      W_g[13,34] := -0.05300187;
      W_g[13,35] := -0.05293896;
      W_g[13,36] := 0.09086524;
      W_g[13,37] := 0.02082952;
      W_g[13,38] := -0.06235110;
      W_g[13,39] := 0.00900952;
      W_g[14,0] := -0.11502921;
      W_g[14,1] := -0.07562436;
      W_g[14,2] := 0.11307055;
      W_g[14,3] := -0.26701322;
      W_g[14,4] := -0.58367014;
      W_g[14,5] := -0.36228108;
      W_g[14,6] := -0.67209059;
      W_g[14,7] := -0.12579566;
      W_g[14,8] := 0.09378675;
      W_g[14,9] := 0.05906596;
      W_g[14,10] := 0.16357109;
      W_g[14,11] := -0.32748589;
      W_g[14,12] := 0.37227204;
      W_g[14,13] := -0.05649122;
      W_g[14,14] := -0.05130398;
      W_g[14,15] := 0.17849237;
      W_g[14,16] := -0.01951551;
      W_g[14,17] := -0.03428079;
      W_g[14,18] := 0.00277206;
      W_g[14,19] := -0.03570505;
      W_g[14,20] := -0.25614583;
      W_g[14,21] := 0.05955129;
      W_g[14,22] := 0.00051241;
      W_g[14,23] := -0.01442853;
      W_g[14,24] := 0.26009023;
      W_g[14,25] := 0.06896590;
      W_g[14,26] := -0.08565364;
      W_g[14,27] := -0.03922650;
      W_g[14,28] := 0.49202508;
      W_g[14,29] := -0.49808294;
      W_g[14,30] := 0.13317353;
      W_g[14,31] := -0.11772110;
      W_g[14,32] := -0.11562508;
      W_g[14,33] := -0.08904682;
      W_g[14,34] := -0.06742100;
      W_g[14,35] := 0.08811268;
      W_g[14,36] := 0.09177279;
      W_g[14,37] := 0.04189566;
      W_g[14,38] := -0.02056031;
      W_g[14,39] := 0.12051180;
      W_g[15,0] := 0.15540718;
      W_g[15,1] := 0.07573265;
      W_g[15,2] := -0.25493059;
      W_g[15,3] := -0.14080612;
      W_g[15,4] := -0.16169477;
      W_g[15,5] := -0.00757927;
      W_g[15,6] := 0.08066899;
      W_g[15,7] := 0.01200249;
      W_g[15,8] := 0.03001926;
      W_g[15,9] := 0.11639266;
      W_g[15,10] := 0.07306892;
      W_g[15,11] := 0.28355977;
      W_g[15,12] := 0.48124212;
      W_g[15,13] := -0.12040935;
      W_g[15,14] := 0.02596140;
      W_g[15,15] := -0.21398795;
      W_g[15,16] := -0.09279459;
      W_g[15,17] := 0.00674920;
      W_g[15,18] := 0.21276073;
      W_g[15,19] := -0.03845788;
      W_g[15,20] := -0.04765760;
      W_g[15,21] := 0.01264688;
      W_g[15,22] := -0.01257103;
      W_g[15,23] := -0.06903563;
      W_g[15,24] := -0.15318221;
      W_g[15,25] := -0.25217903;
      W_g[15,26] := -0.03703345;
      W_g[15,27] := -0.10722972;
      W_g[15,28] := 0.05285160;
      W_g[15,29] := 0.08407086;
      W_g[15,30] := -0.01538745;
      W_g[15,31] := 0.00114667;
      W_g[15,32] := -0.07507251;
      W_g[15,33] := -0.06782222;
      W_g[15,34] := -0.36006817;
      W_g[15,35] := -0.05444269;
      W_g[15,36] := -0.01375175;
      W_g[15,37] := -0.02703385;
      W_g[15,38] := 0.45141658;
      W_g[15,39] := -0.03576548;
      W_g[16,0] := -0.01573141;
      W_g[16,1] := -0.01249725;
      W_g[16,2] := -0.01918053;
      W_g[16,3] := -0.32394302;
      W_g[16,4] := -0.06679904;
      W_g[16,5] := 0.09351813;
      W_g[16,6] := -0.03767738;
      W_g[16,7] := 0.01552502;
      W_g[16,8] := 0.02639228;
      W_g[16,9] := 0.27829525;
      W_g[16,10] := 0.01795475;
      W_g[16,11] := 0.61483020;
      W_g[16,12] := -0.23530579;
      W_g[16,13] := -0.10427370;
      W_g[16,14] := -0.00830992;
      W_g[16,15] := -0.04126130;
      W_g[16,16] := 0.02147032;
      W_g[16,17] := 0.22274575;
      W_g[16,18] := -0.05346655;
      W_g[16,19] := 0.59863454;
      W_g[16,20] := 0.02781765;
      W_g[16,21] := 0.03784034;
      W_g[16,22] := -0.01627534;
      W_g[16,23] := -0.09212849;
      W_g[16,24] := 0.20988049;
      W_g[16,25] := 0.11980043;
      W_g[16,26] := -0.06347527;
      W_g[16,27] := 0.03875433;
      W_g[16,28] := -0.00814277;
      W_g[16,29] := -0.01749807;
      W_g[16,30] := -0.11471809;
      W_g[16,31] := 0.03057062;
      W_g[16,32] := 0.05926932;
      W_g[16,33] := 0.07752163;
      W_g[16,34] := 0.30541685;
      W_g[16,35] := 0.08390119;
      W_g[16,36] := 0.01792176;
      W_g[16,37] := 0.07683819;
      W_g[16,38] := -0.12264256;
      W_g[16,39] := -0.29801413;
      W_g[17,0] := -0.20019235;
      W_g[17,1] := 0.08634444;
      W_g[17,2] := 0.35990810;
      W_g[17,3] := -0.54319084;
      W_g[17,4] := 0.10491174;
      W_g[17,5] := -0.24461722;
      W_g[17,6] := 0.00542844;
      W_g[17,7] := -0.00443292;
      W_g[17,8] := -0.13760753;
      W_g[17,9] := 0.17179628;
      W_g[17,10] := 0.57468456;
      W_g[17,11] := 0.84765750;
      W_g[17,12] := -0.84660238;
      W_g[17,13] := -0.02827467;
      W_g[17,14] := 0.09285270;
      W_g[17,15] := 0.00605520;
      W_g[17,16] := -0.23755617;
      W_g[17,17] := 0.01386433;
      W_g[17,18] := 0.00373611;
      W_g[17,19] := 0.64604604;
      W_g[17,20] := -0.30180034;
      W_g[17,21] := -0.71723890;
      W_g[17,22] := -0.23780504;
      W_g[17,23] := 0.04141965;
      W_g[17,24] := -0.74509096;
      W_g[17,25] := -0.75259161;
      W_g[17,26] := 0.24358149;
      W_g[17,27] := 0.62698990;
      W_g[17,28] := -0.24088508;
      W_g[17,29] := 0.06953070;
      W_g[17,30] := -0.33534220;
      W_g[17,31] := -0.02631341;
      W_g[17,32] := -0.30826521;
      W_g[17,33] := -0.45180380;
      W_g[17,34] := -0.90610892;
      W_g[17,35] := -0.06815604;
      W_g[17,36] := -0.14631121;
      W_g[17,37] := 0.17388295;
      W_g[17,38] := 0.13864316;
      W_g[17,39] := 0.17807765;
      W_g[18,0] := -0.46607670;
      W_g[18,1] := 0.10845635;
      W_g[18,2] := 0.22516194;
      W_g[18,3] := 0.30607522;
      W_g[18,4] := -0.15093884;
      W_g[18,5] := 0.01696070;
      W_g[18,6] := 0.16042185;
      W_g[18,7] := -0.10679442;
      W_g[18,8] := 0.20514138;
      W_g[18,9] := -0.13397862;
      W_g[18,10] := 0.02242056;
      W_g[18,11] := -0.19990624;
      W_g[18,12] := 0.38241696;
      W_g[18,13] := -0.01298471;
      W_g[18,14] := -0.00218331;
      W_g[18,15] := -0.04433896;
      W_g[18,16] := -0.26164895;
      W_g[18,17] := 0.05559360;
      W_g[18,18] := -0.06075819;
      W_g[18,19] := -0.05308994;
      W_g[18,20] := -0.13432083;
      W_g[18,21] := -0.33185339;
      W_g[18,22] := -0.08431048;
      W_g[18,23] := -0.16004905;
      W_g[18,24] := -0.36850065;
      W_g[18,25] := -0.04567018;
      W_g[18,26] := -0.34792730;
      W_g[18,27] := -0.06563149;
      W_g[18,28] := 0.04670760;
      W_g[18,29] := 0.06350503;
      W_g[18,30] := -0.07850740;
      W_g[18,31] := 0.16866533;
      W_g[18,32] := 0.02046569;
      W_g[18,33] := 0.05549860;
      W_g[18,34] := 0.01890240;
      W_g[18,35] := -0.02811935;
      W_g[18,36] := 0.03381456;
      W_g[18,37] := 0.11580943;
      W_g[18,38] := -0.11624962;
      W_g[18,39] := -0.03905239;
      W_g[19,0] := 0.01773376;
      W_g[19,1] := -0.05072702;
      W_g[19,2] := -0.00225121;
      W_g[19,3] := -0.01785041;
      W_g[19,4] := 0.04858205;
      W_g[19,5] := -0.01839915;
      W_g[19,6] := -0.04408873;
      W_g[19,7] := -0.01353623;
      W_g[19,8] := -0.00090088;
      W_g[19,9] := -0.00116132;
      W_g[19,10] := 0.00882178;
      W_g[19,11] := -0.03854829;
      W_g[19,12] := 0.03738030;
      W_g[19,13] := -0.01948604;
      W_g[19,14] := -0.45808697;
      W_g[19,15] := -0.26110804;
      W_g[19,16] := 0.00333187;
      W_g[19,17] := -0.25176817;
      W_g[19,18] := 0.08445162;
      W_g[19,19] := 0.26523203;
      W_g[19,20] := -0.05709776;
      W_g[19,21] := -0.05241840;
      W_g[19,22] := 0.01751016;
      W_g[19,23] := -0.00974986;
      W_g[19,24] := 0.27344036;
      W_g[19,25] := 0.32422283;
      W_g[19,26] := -0.04881701;
      W_g[19,27] := -0.02297378;
      W_g[19,28] := -0.06826914;
      W_g[19,29] := -0.11992263;
      W_g[19,30] := 0.01903425;
      W_g[19,31] := 0.02200578;
      W_g[19,32] := -0.04815840;
      W_g[19,33] := -0.11233919;
      W_g[19,34] := -0.23930897;
      W_g[19,35] := 0.02726550;
      W_g[19,36] := -0.00201288;
      W_g[19,37] := 0.05262006;
      W_g[19,38] := -0.04631574;
      W_g[19,39] := -0.25027138;
      W_g[20,0] := -0.17776611;
      W_g[20,1] := -0.49992636;
      W_g[20,2] := 0.03143674;
      W_g[20,3] := 0.15612000;
      W_g[20,4] := -0.50436848;
      W_g[20,5] := 0.02739897;
      W_g[20,6] := -0.10362915;
      W_g[20,7] := 0.35108495;
      W_g[20,8] := 0.19622006;
      W_g[20,9] := 0.38027030;
      W_g[20,10] := -0.53794569;
      W_g[20,11] := 0.05582263;
      W_g[20,12] := -0.17187732;
      W_g[20,13] := -0.14350507;
      W_g[20,14] := 0.04435784;
      W_g[20,15] := -0.00301744;
      W_g[20,16] := 0.05593058;
      W_g[20,17] := 0.00574902;
      W_g[20,18] := 0.02816820;
      W_g[20,19] := -0.00896498;
      W_g[20,20] := -0.27302650;
      W_g[20,21] := -0.10916554;
      W_g[20,22] := 0.07598325;
      W_g[20,23] := 0.07597133;
      W_g[20,24] := -0.20816125;
      W_g[20,25] := -0.00556583;
      W_g[20,26] := 0.15926160;
      W_g[20,27] := 0.04909170;
      W_g[20,28] := -0.30622017;
      W_g[20,29] := 0.16263185;
      W_g[20,30] := 0.06980544;
      W_g[20,31] := 0.18102454;
      W_g[20,32] := 0.01593671;
      W_g[20,33] := -0.04853294;
      W_g[20,34] := -0.09243315;
      W_g[20,35] := 0.03795157;
      W_g[20,36] := -0.01642190;
      W_g[20,37] := 0.06450415;
      W_g[20,38] := -0.01715147;
      W_g[20,39] := -0.05797761;
      W_g[21,0] := 0.04719520;
      W_g[21,1] := 0.01569074;
      W_g[21,2] := -0.00857600;
      W_g[21,3] := 0.36854166;
      W_g[21,4] := -0.29962948;
      W_g[21,5] := 0.11101421;
      W_g[21,6] := -0.14704654;
      W_g[21,7] := -0.25060529;
      W_g[21,8] := 0.03979661;
      W_g[21,9] := -0.37424278;
      W_g[21,10] := 0.33715650;
      W_g[21,11] := 0.20566781;
      W_g[21,12] := -0.55089366;
      W_g[21,13] := -0.34874550;
      W_g[21,14] := -0.00000745;
      W_g[21,15] := 0.11779826;
      W_g[21,16] := -0.01198818;
      W_g[21,17] := -0.09557019;
      W_g[21,18] := -0.38575107;
      W_g[21,19] := 0.10345905;
      W_g[21,20] := 0.17967871;
      W_g[21,21] := -0.02546586;
      W_g[21,22] := 0.02202458;
      W_g[21,23] := -0.47533408;
      W_g[21,24] := -0.07804859;
      W_g[21,25] := -0.20474817;
      W_g[21,26] := 0.09593988;
      W_g[21,27] := -0.20002005;
      W_g[21,28] := 0.14636038;
      W_g[21,29] := 0.27730727;
      W_g[21,30] := 0.03117772;
      W_g[21,31] := 0.06990665;
      W_g[21,32] := 0.05139569;
      W_g[21,33] := 0.08534111;
      W_g[21,34] := 0.34672982;
      W_g[21,35] := 0.01232039;
      W_g[21,36] := -0.05206082;
      W_g[21,37] := -0.01625307;
      W_g[21,38] := 0.20143867;
      W_g[21,39] := -0.10067950;
      W_g[22,0] := 0.11665134;
      W_g[22,1] := 0.10529415;
      W_g[22,2] := 0.22086281;
      W_g[22,3] := -0.12558044;
      W_g[22,4] := -0.00237558;
      W_g[22,5] := 0.19240804;
      W_g[22,6] := -0.24772990;
      W_g[22,7] := 0.08354132;
      W_g[22,8] := -0.20447712;
      W_g[22,9] := 0.03358927;
      W_g[22,10] := -0.15093991;
      W_g[22,11] := -0.03152904;
      W_g[22,12] := 0.23958053;
      W_g[22,13] := -0.10689051;
      W_g[22,14] := 0.14513183;
      W_g[22,15] := 0.20699252;
      W_g[22,16] := -0.00007249;
      W_g[22,17] := 0.01122855;
      W_g[22,18] := -0.00866538;
      W_g[22,19] := 0.10550721;
      W_g[22,20] := -0.14577182;
      W_g[22,21] := 0.25070757;
      W_g[22,22] := 0.07765597;
      W_g[22,23] := 0.12089684;
      W_g[22,24] := 0.42342681;
      W_g[22,25] := 0.12979737;
      W_g[22,26] := 0.16623591;
      W_g[22,27] := -0.09820254;
      W_g[22,28] := 0.03250218;
      W_g[22,29] := 0.11340379;
      W_g[22,30] := 0.08371338;
      W_g[22,31] := 0.10858538;
      W_g[22,32] := -0.09717516;
      W_g[22,33] := -0.05043048;
      W_g[22,34] := -0.12874730;
      W_g[22,35] := -0.16679265;
      W_g[22,36] := 0.06777173;
      W_g[22,37] := -0.19872338;
      W_g[22,38] := -0.09894791;
      W_g[22,39] := -0.29871914;
      W_g[23,0] := -0.07641292;
      W_g[23,1] := -0.00534786;
      W_g[23,2] := 0.20778368;
      W_g[23,3] := 0.22361241;
      W_g[23,4] := 0.03807362;
      W_g[23,5] := -0.02697703;
      W_g[23,6] := -0.13366827;
      W_g[23,7] := -0.03372496;
      W_g[23,8] := -0.11303925;
      W_g[23,9] := -0.14616819;
      W_g[23,10] := 0.00094925;
      W_g[23,11] := 0.17858963;
      W_g[23,12] := -0.02489791;
      W_g[23,13] := -0.03910236;
      W_g[23,14] := -0.02416698;
      W_g[23,15] := -0.25673768;
      W_g[23,16] := 0.30395365;
      W_g[23,17] := -0.01390388;
      W_g[23,18] := 0.00377696;
      W_g[23,19] := 0.08999401;
      W_g[23,20] := -0.40618902;
      W_g[23,21] := -0.18011197;
      W_g[23,22] := -0.10348500;
      W_g[23,23] := 0.01184078;
      W_g[23,24] := -0.60941619;
      W_g[23,25] := -0.17570031;
      W_g[23,26] := 0.09114521;
      W_g[23,27] := 0.07809471;
      W_g[23,28] := -0.03781823;
      W_g[23,29] := -0.02985572;
      W_g[23,30] := -0.10175200;
      W_g[23,31] := 0.07091261;
      W_g[23,32] := 0.00975894;
      W_g[23,33] := 0.07413130;
      W_g[23,34] := 0.04860087;
      W_g[23,35] := -0.06112134;
      W_g[23,36] := -0.01834961;
      W_g[23,37] := -0.06767160;
      W_g[23,38] := 0.04615815;
      W_g[23,39] := 0.03219241;
      W_g[24,0] := 0.14109130;
      W_g[24,1] := 0.23656085;
      W_g[24,2] := -0.05220996;
      W_g[24,3] := -0.08191337;
      W_g[24,4] := -0.59643692;
      W_g[24,5] := -0.08740985;
      W_g[24,6] := 0.51112539;
      W_g[24,7] := -0.08679886;
      W_g[24,8] := -0.03170026;
      W_g[24,9] := -0.04040290;
      W_g[24,10] := 0.42674446;
      W_g[24,11] := 0.22892350;
      W_g[24,12] := 0.06517982;
      W_g[24,13] := -0.07052775;
      W_g[24,14] := 0.00610844;
      W_g[24,15] := -0.14473575;
      W_g[24,16] := 0.11628936;
      W_g[24,17] := 0.00950560;
      W_g[24,18] := -0.05220868;
      W_g[24,19] := -0.21057445;
      W_g[24,20] := 0.15953180;
      W_g[24,21] := 0.03443460;
      W_g[24,22] := 0.02498991;
      W_g[24,23] := 0.15479933;
      W_g[24,24] := 0.31532544;
      W_g[24,25] := -0.07248386;
      W_g[24,26] := 0.22804081;
      W_g[24,27] := -0.23870072;
      W_g[24,28] := 0.07509667;
      W_g[24,29] := -0.04223498;
      W_g[24,30] := 0.02754644;
      W_g[24,31] := 0.04945280;
      W_g[24,32] := -0.12835518;
      W_g[24,33] := -0.16013861;
      W_g[24,34] := -0.20117347;
      W_g[24,35] := -0.09332737;
      W_g[24,36] := -0.27658218;
      W_g[24,37] := -0.14927265;
      W_g[24,38] := -0.28982732;
      W_g[24,39] := 0.01216547;
      W_g[25,0] := 0.00249727;
      W_g[25,1] := 0.02321395;
      W_g[25,2] := 0.03579676;
      W_g[25,3] := -0.32325658;
      W_g[25,4] := 0.07457885;
      W_g[25,5] := 0.01599968;
      W_g[25,6] := -0.19957243;
      W_g[25,7] := 0.12909044;
      W_g[25,8] := 0.00623424;
      W_g[25,9] := 0.26816839;
      W_g[25,10] := -0.23799382;
      W_g[25,11] := -0.18556090;
      W_g[25,12] := -0.03897551;
      W_g[25,13] := -0.07030228;
      W_g[25,14] := -0.06287792;
      W_g[25,15] := 0.17744720;
      W_g[25,16] := -0.03842967;
      W_g[25,17] := -0.06559484;
      W_g[25,18] := 0.02993315;
      W_g[25,19] := 0.08945196;
      W_g[25,20] := -0.00580116;
      W_g[25,21] := -0.02753790;
      W_g[25,22] := -0.02607165;
      W_g[25,23] := -0.00466925;
      W_g[25,24] := -0.84821171;
      W_g[25,25] := 0.23694646;
      W_g[25,26] := -0.14543480;
      W_g[25,27] := -0.15780894;
      W_g[25,28] := -0.27692312;
      W_g[25,29] := -0.04585484;
      W_g[25,30] := -0.03756009;
      W_g[25,31] := -0.08991528;
      W_g[25,32] := 0.00971850;
      W_g[25,33] := 0.08656777;
      W_g[25,34] := 0.12360313;
      W_g[25,35] := -0.08704287;
      W_g[25,36] := -0.50061452;
      W_g[25,37] := 0.06715164;
      W_g[25,38] := 0.03072628;
      W_g[25,39] := -0.05923472;
      W_g[26,0] := 0.19895676;
      W_g[26,1] := 0.01795273;
      W_g[26,2] := -0.08949947;
      W_g[26,3] := -0.06816271;
      W_g[26,4] := -0.12828159;
      W_g[26,5] := 0.00080027;
      W_g[26,6] := 0.16275345;
      W_g[26,7] := 0.14247812;
      W_g[26,8] := -0.05336298;
      W_g[26,9] := 0.16001105;
      W_g[26,10] := -0.00170321;
      W_g[26,11] := -0.10854331;
      W_g[26,12] := 0.11391646;
      W_g[26,13] := 0.31833315;
      W_g[26,14] := -0.00052231;
      W_g[26,15] := 0.04305906;
      W_g[26,16] := -0.00767927;
      W_g[26,17] := -0.03174791;
      W_g[26,18] := -1.20069015;
      W_g[26,19] := 0.08255526;
      W_g[26,20] := -0.47470504;
      W_g[26,21] := 0.21856050;
      W_g[26,22] := 0.04315476;
      W_g[26,23] := 0.15731587;
      W_g[26,24] := -0.16662689;
      W_g[26,25] := -0.36638814;
      W_g[26,26] := -0.28305781;
      W_g[26,27] := -0.09379881;
      W_g[26,28] := -0.24579851;
      W_g[26,29] := 0.01016386;
      W_g[26,30] := 0.01751088;
      W_g[26,31] := 0.15965039;
      W_g[26,32] := 0.00510592;
      W_g[26,33] := 0.09451680;
      W_g[26,34] := 0.02374958;
      W_g[26,35] := -0.10228859;
      W_g[26,36] := 0.04589900;
      W_g[26,37] := -0.01942009;
      W_g[26,38] := 0.15447062;
      W_g[26,39] := -0.00123656;
      W_g[27,0] := -0.14282966;
      W_g[27,1] := 0.03789151;
      W_g[27,2] := 0.02735430;
      W_g[27,3] := -0.02859589;
      W_g[27,4] := 0.11969381;
      W_g[27,5] := -0.08108735;
      W_g[27,6] := -0.48059788;
      W_g[27,7] := 0.11670560;
      W_g[27,8] := 0.02436283;
      W_g[27,9] := 0.15240525;
      W_g[27,10] := 0.60784400;
      W_g[27,11] := 0.16673699;
      W_g[27,12] := -0.11131126;
      W_g[27,13] := 0.39158168;
      W_g[27,14] := -0.01387984;
      W_g[27,15] := 0.03263223;
      W_g[27,16] := 0.07995110;
      W_g[27,17] := -0.01656702;
      W_g[27,18] := 0.16666247;
      W_g[27,19] := -0.07363571;
      W_g[27,20] := -0.26380217;
      W_g[27,21] := 0.36762938;
      W_g[27,22] := 0.10293096;
      W_g[27,23] := -0.21954748;
      W_g[27,24] := -0.19905801;
      W_g[27,25] := 0.00590560;
      W_g[27,26] := -0.07474038;
      W_g[27,27] := -0.00682373;
      W_g[27,28] := 0.00600550;
      W_g[27,29] := 0.52201474;
      W_g[27,30] := 0.10763236;
      W_g[27,31] := 0.20513408;
      W_g[27,32] := 0.08530629;
      W_g[27,33] := 0.18354966;
      W_g[27,34] := 0.20833531;
      W_g[27,35] := -0.02688346;
      W_g[27,36] := -0.05211073;
      W_g[27,37] := -0.10546255;
      W_g[27,38] := -0.16810939;
      W_g[27,39] := 0.04055268;
      W_g[28,0] := -0.12039233;
      W_g[28,1] := 0.03123983;
      W_g[28,2] := -0.28947538;
      W_g[28,3] := -0.24017365;
      W_g[28,4] := 0.29521075;
      W_g[28,5] := 0.08690419;
      W_g[28,6] := 0.01901748;
      W_g[28,7] := -0.23417597;
      W_g[28,8] := 0.43286511;
      W_g[28,9] := 0.02607675;
      W_g[28,10] := 0.19849846;
      W_g[28,11] := -0.06265938;
      W_g[28,12] := 0.09416307;
      W_g[28,13] := -0.05105516;
      W_g[28,14] := -0.01597860;
      W_g[28,15] := 0.14792809;
      W_g[28,16] := 0.14414477;
      W_g[28,17] := -0.02288275;
      W_g[28,18] := -0.03377746;
      W_g[28,19] := -0.15792006;
      W_g[28,20] := -0.21533181;
      W_g[28,21] := 0.08094171;
      W_g[28,22] := 0.00793070;
      W_g[28,23] := 0.03326877;
      W_g[28,24] := 0.04408788;
      W_g[28,25] := -0.11347675;
      W_g[28,26] := 0.14422546;
      W_g[28,27] := 0.19584695;
      W_g[28,28] := -0.13756958;
      W_g[28,29] := -0.12223729;
      W_g[28,30] := 0.02110463;
      W_g[28,31] := 0.03519979;
      W_g[28,32] := -0.05562153;
      W_g[28,33] := -0.06591920;
      W_g[28,34] := 0.04866378;
      W_g[28,35] := -0.09032071;
      W_g[28,36] := 0.03939996;
      W_g[28,37] := -0.08595932;
      W_g[28,38] := 0.01556356;
      W_g[28,39] := -0.17334549;
      W_g[29,0] := -0.01603005;
      W_g[29,1] := 0.00894765;
      W_g[29,2] := 0.04728428;
      W_g[29,3] := 0.13398947;
      W_g[29,4] := -0.08206625;
      W_g[29,5] := 0.43515241;
      W_g[29,6] := -0.08524376;
      W_g[29,7] := 0.12636763;
      W_g[29,8] := -0.07064829;
      W_g[29,9] := 0.02922662;
      W_g[29,10] := 0.16617142;
      W_g[29,11] := -0.03181689;
      W_g[29,12] := -0.18755385;
      W_g[29,13] := 0.04736114;
      W_g[29,14] := 0.00172536;
      W_g[29,15] := 0.02388163;
      W_g[29,16] := -0.00605842;
      W_g[29,17] := -0.00226685;
      W_g[29,18] := 0.18417786;
      W_g[29,19] := 0.02931385;
      W_g[29,20] := -0.10084365;
      W_g[29,21] := -0.03299641;
      W_g[29,22] := -0.00275616;
      W_g[29,23] := 0.02141913;
      W_g[29,24] := 0.00477037;
      W_g[29,25] := 0.05081034;
      W_g[29,26] := -0.19006838;
      W_g[29,27] := -0.14232871;
      W_g[29,28] := 0.06605857;
      W_g[29,29] := -0.26251897;
      W_g[29,30] := -0.00548652;
      W_g[29,31] := 0.03245487;
      W_g[29,32] := -0.05614575;
      W_g[29,33] := -0.08672421;
      W_g[29,34] := -0.19275941;
      W_g[29,35] := -0.02231585;
      W_g[29,36] := 0.00673404;
      W_g[29,37] := -0.02077745;
      W_g[29,38] := 0.02013531;
      W_g[29,39] := 0.21206558;
      W_g[30,0] := 0.06752372;
      W_g[30,1] := 0.04914160;
      W_g[30,2] := 0.03581399;
      W_g[30,3] := 0.55463815;
      W_g[30,4] := 0.19955039;
      W_g[30,5] := -0.29638356;
      W_g[30,6] := 0.61677969;
      W_g[30,7] := -0.08204620;
      W_g[30,8] := -0.02945163;
      W_g[30,9] := -0.33782583;
      W_g[30,10] := 0.03250416;
      W_g[30,11] := 0.32107306;
      W_g[30,12] := 0.06659118;
      W_g[30,13] := 0.29332143;
      W_g[30,14] := -0.02582538;
      W_g[30,15] := 0.62199312;
      W_g[30,16] := 0.28212488;
      W_g[30,17] := -0.23582231;
      W_g[30,18] := 0.33779177;
      W_g[30,19] := 0.50508004;
      W_g[30,20] := -0.04146927;
      W_g[30,21] := 0.00146027;
      W_g[30,22] := 0.10298456;
      W_g[30,23] := -0.13510256;
      W_g[30,24] := 0.08098176;
      W_g[30,25] := -0.07603540;
      W_g[30,26] := 0.11315724;
      W_g[30,27] := 0.12087354;
      W_g[30,28] := -0.23194072;
      W_g[30,29] := 0.06172852;
      W_g[30,30] := 0.06911052;
      W_g[30,31] := 0.33844078;
      W_g[30,32] := 0.07554214;
      W_g[30,33] := 0.01718852;
      W_g[30,34] := -0.07873586;
      W_g[30,35] := -0.07006503;
      W_g[30,36] := 0.00541107;
      W_g[30,37] := -0.08336300;
      W_g[30,38] := 0.02301235;
      W_g[30,39] := 0.23563193;
      W_g[31,0] := 0.18860947;
      W_g[31,1] := -0.02123935;
      W_g[31,2] := -0.26690537;
      W_g[31,3] := 0.12378932;
      W_g[31,4] := 0.09037927;
      W_g[31,5] := -0.03088225;
      W_g[31,6] := -0.17878367;
      W_g[31,7] := 0.02112429;
      W_g[31,8] := 0.03763676;
      W_g[31,9] := -0.02504454;
      W_g[31,10] := -0.01659736;
      W_g[31,11] := 0.16001292;
      W_g[31,12] := -0.06862063;
      W_g[31,13] := -0.08124028;
      W_g[31,14] := -0.00468529;
      W_g[31,15] := -0.14859970;
      W_g[31,16] := -0.30615747;
      W_g[31,17] := -0.02353984;
      W_g[31,18] := 0.01195374;
      W_g[31,19] := 0.04420421;
      W_g[31,20] := -0.08521901;
      W_g[31,21] := 0.06032958;
      W_g[31,22] := 0.01825500;
      W_g[31,23] := 0.05283485;
      W_g[31,24] := -0.25803921;
      W_g[31,25] := 0.03302622;
      W_g[31,26] := 0.16146830;
      W_g[31,27] := 0.17279540;
      W_g[31,28] := 0.01809685;
      W_g[31,29] := 0.02630481;
      W_g[31,30] := 0.03338469;
      W_g[31,31] := 0.45954949;
      W_g[31,32] := -0.04697010;
      W_g[31,33] := 0.03801997;
      W_g[31,34] := 0.22326140;
      W_g[31,35] := -0.18952455;
      W_g[31,36] := 0.00136513;
      W_g[31,37] := -0.27123162;
      W_g[31,38] := -0.07247190;
      W_g[31,39] := 0.23167513;
      W_o[0,0] := 0.42249125;
      W_o[0,1] := -0.64850706;
      W_o[0,2] := -0.08193821;
      W_o[0,3] := -0.33892727;
      W_o[0,4] := 0.05321682;
      W_o[0,5] := 0.11530717;
      W_o[0,6] := 0.32608813;
      W_o[0,7] := -0.13539509;
      W_o[0,8] := 0.20117587;
      W_o[0,9] := -0.31878343;
      W_o[0,10] := -0.17219098;
      W_o[0,11] := 0.14882079;
      W_o[0,12] := 0.11313346;
      W_o[0,13] := -0.10760950;
      W_o[0,14] := 0.01743469;
      W_o[0,15] := 0.01349122;
      W_o[0,16] := -0.01363511;
      W_o[0,17] := -0.00418937;
      W_o[0,18] := -0.08654208;
      W_o[0,19] := 0.01018774;
      W_o[0,20] := 0.37044030;
      W_o[0,21] := 0.87406963;
      W_o[0,22] := 0.05330493;
      W_o[0,23] := -0.60551524;
      W_o[0,24] := 0.00528000;
      W_o[0,25] := 0.00492091;
      W_o[0,26] := -0.73618817;
      W_o[0,27] := 0.86269325;
      W_o[0,28] := 0.67136478;
      W_o[0,29] := -0.14723247;
      W_o[0,30] := -0.17640491;
      W_o[0,31] := 0.00200789;
      W_o[0,32] := -0.11784527;
      W_o[0,33] := 0.32575944;
      W_o[0,34] := 0.11160263;
      W_o[0,35] := -0.05652209;
      W_o[0,36] := 0.04402122;
      W_o[0,37] := 0.08225929;
      W_o[0,38] := 0.20138605;
      W_o[0,39] := -0.07881875;
      W_o[1,0] := -1.27534890;
      W_o[1,1] := -0.27924889;
      W_o[1,2] := -0.75771481;
      W_o[1,3] := -0.18380418;
      W_o[1,4] := -0.39482769;
      W_o[1,5] := 0.10104305;
      W_o[1,6] := -0.34825188;
      W_o[1,7] := -0.63163066;
      W_o[1,8] := -1.08178067;
      W_o[1,9] := -0.97093791;
      W_o[1,10] := -0.20904520;
      W_o[1,11] := -0.29529026;
      W_o[1,12] := -0.14393961;
      W_o[1,13] := -0.01520389;
      W_o[1,14] := 0.00541295;
      W_o[1,15] := -0.02735653;
      W_o[1,16] := -0.07699423;
      W_o[1,17] := 0.08873669;
      W_o[1,18] := 0.18124166;
      W_o[1,19] := -0.01098941;
      W_o[1,20] := 0.13787243;
      W_o[1,21] := 0.26410136;
      W_o[1,22] := 0.06537609;
      W_o[1,23] := -0.15175536;
      W_o[1,24] := -0.11301857;
      W_o[1,25] := -0.10047740;
      W_o[1,26] := 0.11024941;
      W_o[1,27] := 0.24368817;
      W_o[1,28] := 0.59257942;
      W_o[1,29] := 0.02251752;
      W_o[1,30] := 0.20542605;
      W_o[1,31] := 0.05349508;
      W_o[1,32] := 0.07199062;
      W_o[1,33] := 0.06075877;
      W_o[1,34] := 0.17365526;
      W_o[1,35] := -0.04894430;
      W_o[1,36] := -0.02975028;
      W_o[1,37] := -0.12903002;
      W_o[1,38] := 0.08992038;
      W_o[1,39] := 0.10337646;
      W_o[2,0] := 0.30405313;
      W_o[2,1] := 0.00766394;
      W_o[2,2] := -0.18612629;
      W_o[2,3] := 0.15926282;
      W_o[2,4] := 0.50370109;
      W_o[2,5] := 0.69898289;
      W_o[2,6] := 1.03120697;
      W_o[2,7] := 0.06395171;
      W_o[2,8] := 0.13832410;
      W_o[2,9] := 0.10960636;
      W_o[2,10] := -0.42085138;
      W_o[2,11] := 0.39040789;
      W_o[2,12] := 0.06325981;
      W_o[2,13] := 0.40687191;
      W_o[2,14] := 0.04082680;
      W_o[2,15] := -0.00324509;
      W_o[2,16] := 0.01833900;
      W_o[2,17] := 0.11513314;
      W_o[2,18] := 0.12066066;
      W_o[2,19] := 0.01082493;
      W_o[2,20] := -0.16976321;
      W_o[2,21] := 0.53049803;
      W_o[2,22] := 0.15725319;
      W_o[2,23] := -0.34637845;
      W_o[2,24] := 1.58245826;
      W_o[2,25] := 1.47554839;
      W_o[2,26] := -0.00448998;
      W_o[2,27] := 0.14077175;
      W_o[2,28] := -0.37107602;
      W_o[2,29] := 0.02695022;
      W_o[2,30] := 0.19601339;
      W_o[2,31] := 0.17389217;
      W_o[2,32] := 0.14344938;
      W_o[2,33] := 0.81406116;
      W_o[2,34] := 1.72799015;
      W_o[2,35] := -0.12091801;
      W_o[2,36] := 0.16224357;
      W_o[2,37] := -0.33939198;
      W_o[2,38] := 0.05670876;
      W_o[2,39] := 0.09963638;
      W_o[3,0] := -0.26549935;
      W_o[3,1] := -0.11039463;
      W_o[3,2] := -0.37164780;
      W_o[3,3] := 0.15892562;
      W_o[3,4] := -0.06230325;
      W_o[3,5] := -0.37457275;
      W_o[3,6] := 0.24259707;
      W_o[3,7] := 0.37691608;
      W_o[3,8] := -0.42493910;
      W_o[3,9] := 0.27702668;
      W_o[3,10] := 0.36755127;
      W_o[3,11] := -0.49238053;
      W_o[3,12] := -0.28828865;
      W_o[3,13] := -0.19150881;
      W_o[3,14] := -0.67414224;
      W_o[3,15] := -0.02529657;
      W_o[3,16] := 0.29622570;
      W_o[3,17] := 0.45850250;
      W_o[3,18] := 0.04778790;
      W_o[3,19] := 0.51993376;
      W_o[3,20] := -0.20207447;
      W_o[3,21] := 0.18979242;
      W_o[3,22] := -0.07848933;
      W_o[3,23] := -0.01705214;
      W_o[3,24] := 0.01806957;
      W_o[3,25] := 0.02297689;
      W_o[3,26] := -0.01870384;
      W_o[3,27] := -0.17662346;
      W_o[3,28] := -0.04692467;
      W_o[3,29] := -0.17209335;
      W_o[3,30] := -0.24459122;
      W_o[3,31] := 0.07113735;
      W_o[3,32] := 0.00606646;
      W_o[3,33] := -0.05090882;
      W_o[3,34] := 0.08984744;
      W_o[3,35] := -0.16125588;
      W_o[3,36] := -0.00926951;
      W_o[3,37] := -0.15794532;
      W_o[3,38] := 0.07680272;
      W_o[3,39] := 1.02147377;
      W_o[4,0] := 0.17977053;
      W_o[4,1] := 0.03995879;
      W_o[4,2] := -0.05187562;
      W_o[4,3] := -0.00068046;
      W_o[4,4] := 0.00082433;
      W_o[4,5] := -0.17477073;
      W_o[4,6] := 0.18298250;
      W_o[4,7] := 0.01242155;
      W_o[4,8] := -0.10564039;
      W_o[4,9] := 0.28895974;
      W_o[4,10] := -0.16322204;
      W_o[4,11] := 0.10945952;
      W_o[4,12] := -0.03262473;
      W_o[4,13] := -0.11646359;
      W_o[4,14] := 0.00214941;
      W_o[4,15] := -0.01470709;
      W_o[4,16] := 0.07081575;
      W_o[4,17] := -0.00195280;
      W_o[4,18] := 0.90504497;
      W_o[4,19] := 0.06995305;
      W_o[4,20] := 0.12764473;
      W_o[4,21] := -0.13823217;
      W_o[4,22] := -0.10447618;
      W_o[4,23] := -0.07500455;
      W_o[4,24] := -0.22946472;
      W_o[4,25] := 0.20651680;
      W_o[4,26] := 0.08378618;
      W_o[4,27] := 0.07185337;
      W_o[4,28] := 0.15295289;
      W_o[4,29] := 0.80911016;
      W_o[4,30] := -0.12649418;
      W_o[4,31] := 0.29769754;
      W_o[4,32] := -0.10073072;
      W_o[4,33] := -0.19524801;
      W_o[4,34] := -0.00692285;
      W_o[4,35] := 0.15373145;
      W_o[4,36] := 0.01237739;
      W_o[4,37] := 0.13210568;
      W_o[4,38] := 0.15424773;
      W_o[4,39] := -0.01015362;
      W_o[5,0] := 0.28912961;
      W_o[5,1] := 2.07105112;
      W_o[5,2] := 0.01252856;
      W_o[5,3] := 0.34673738;
      W_o[5,4] := 0.21192910;
      W_o[5,5] := 0.23409151;
      W_o[5,6] := -0.12695056;
      W_o[5,7] := 0.23784913;
      W_o[5,8] := -0.03728350;
      W_o[5,9] := 0.21514873;
      W_o[5,10] := 0.26284939;
      W_o[5,11] := -0.21792066;
      W_o[5,12] := -0.39795417;
      W_o[5,13] := -0.69216830;
      W_o[5,14] := -0.18849657;
      W_o[5,15] := -0.13393024;
      W_o[5,16] := -0.25170875;
      W_o[5,17] := -0.24293463;
      W_o[5,18] := 0.27309209;
      W_o[5,19] := -0.14950365;
      W_o[5,20] := -0.03219712;
      W_o[5,21] := 0.35288468;
      W_o[5,22] := 0.23942992;
      W_o[5,23] := -0.16948508;
      W_o[5,24] := 1.87266624;
      W_o[5,25] := 1.58824658;
      W_o[5,26] := -0.05295049;
      W_o[5,27] := 0.20530860;
      W_o[5,28] := -0.00417454;
      W_o[5,29] := -0.04709773;
      W_o[5,30] := 0.14920191;
      W_o[5,31] := -0.05560581;
      W_o[5,32] := 0.04669352;
      W_o[5,33] := 0.14553502;
      W_o[5,34] := 0.53250414;
      W_o[5,35] := 0.10384236;
      W_o[5,36] := 0.39177659;
      W_o[5,37] := -0.00503783;
      W_o[5,38] := -0.05498653;
      W_o[5,39] := 0.39836636;
      W_o[6,0] := -0.09602387;
      W_o[6,1] := 0.01318664;
      W_o[6,2] := 0.02895827;
      W_o[6,3] := -0.13262498;
      W_o[6,4] := -0.12622669;
      W_o[6,5] := 0.03745453;
      W_o[6,6] := 0.55729073;
      W_o[6,7] := 0.14179020;
      W_o[6,8] := 0.08813037;
      W_o[6,9] := 0.02709752;
      W_o[6,10] := -0.03546845;
      W_o[6,11] := 0.07040328;
      W_o[6,12] := -0.03574698;
      W_o[6,13] := 0.01986431;
      W_o[6,14] := 0.01404128;
      W_o[6,15] := 0.02171072;
      W_o[6,16] := 0.09358315;
      W_o[6,17] := 0.05428468;
      W_o[6,18] := -0.02667183;
      W_o[6,19] := -0.00128908;
      W_o[6,20] := -1.56595874;
      W_o[6,21] := 0.00646133;
      W_o[6,22] := -0.24436766;
      W_o[6,23] := -0.13901594;
      W_o[6,24] := 0.99376416;
      W_o[6,25] := 0.85211402;
      W_o[6,26] := -0.23664802;
      W_o[6,27] := -0.08933339;
      W_o[6,28] := 0.15226653;
      W_o[6,29] := -0.30946207;
      W_o[6,30] := -0.20975208;
      W_o[6,31] := 0.62505847;
      W_o[6,32] := -0.04092027;
      W_o[6,33] := 0.09183368;
      W_o[6,34] := 0.63159341;
      W_o[6,35] := 0.13661051;
      W_o[6,36] := -0.00265529;
      W_o[6,37] := 0.16893734;
      W_o[6,38] := 0.18080245;
      W_o[6,39] := 0.49472585;
      W_o[7,0] := 0.12950280;
      W_o[7,1] := -0.08431699;
      W_o[7,2] := 0.01352446;
      W_o[7,3] := -0.24629471;
      W_o[7,4] := -0.11285538;
      W_o[7,5] := 0.10077246;
      W_o[7,6] := -0.37715051;
      W_o[7,7] := 0.07297357;
      W_o[7,8] := 0.21676154;
      W_o[7,9] := -0.45346865;
      W_o[7,10] := -0.07251467;
      W_o[7,11] := -0.11458308;
      W_o[7,12] := 0.13860887;
      W_o[7,13] := 0.02705087;
      W_o[7,14] := -0.46493185;
      W_o[7,15] := -0.09500964;
      W_o[7,16] := -0.02847600;
      W_o[7,17] := -0.33199629;
      W_o[7,18] := 0.75860929;
      W_o[7,19] := -0.24825610;
      W_o[7,20] := 0.07540248;
      W_o[7,21] := -0.00047477;
      W_o[7,22] := 0.39176366;
      W_o[7,23] := 0.24398798;
      W_o[7,24] := 0.09440543;
      W_o[7,25] := 0.08927973;
      W_o[7,26] := -0.18593012;
      W_o[7,27] := 0.50119442;
      W_o[7,28] := 0.22797424;
      W_o[7,29] := 0.42095158;
      W_o[7,30] := 0.29652157;
      W_o[7,31] := -0.04999515;
      W_o[7,32] := -0.15699139;
      W_o[7,33] := -0.18410453;
      W_o[7,34] := -0.08341311;
      W_o[7,35] := 0.13659917;
      W_o[7,36] := -0.56333482;
      W_o[7,37] := 0.05962496;
      W_o[7,38] := -0.13092983;
      W_o[7,39] := 0.24780601;
      W_o[8,0] := 0.24813814;
      W_o[8,1] := 0.00067703;
      W_o[8,2] := -0.14760867;
      W_o[8,3] := -0.20843014;
      W_o[8,4] := 0.02320351;
      W_o[8,5] := -0.15086000;
      W_o[8,6] := -0.11804635;
      W_o[8,7] := 0.18003957;
      W_o[8,8] := -0.02108677;
      W_o[8,9] := -0.16253571;
      W_o[8,10] := 0.06853176;
      W_o[8,11] := -0.64998335;
      W_o[8,12] := 0.36357620;
      W_o[8,13] := 0.08369323;
      W_o[8,14] := 0.01761020;
      W_o[8,15] := -0.24554460;
      W_o[8,16] := 0.21399209;
      W_o[8,17] := -0.16698237;
      W_o[8,18] := -0.05301695;
      W_o[8,19] := -1.55503678;
      W_o[8,20] := -0.04698478;
      W_o[8,21] := -0.14936455;
      W_o[8,22] := 0.07500248;
      W_o[8,23] := -0.13922599;
      W_o[8,24] := 0.59468526;
      W_o[8,25] := 0.81987101;
      W_o[8,26] := -0.03043681;
      W_o[8,27] := 0.27328554;
      W_o[8,28] := 0.10655938;
      W_o[8,29] := -0.01688519;
      W_o[8,30] := 0.12638046;
      W_o[8,31] := 0.29698491;
      W_o[8,32] := 0.25925279;
      W_o[8,33] := 0.19317611;
      W_o[8,34] := 0.61168981;
      W_o[8,35] := 0.15048993;
      W_o[8,36] := -0.07168282;
      W_o[8,37] := 0.00242552;
      W_o[8,38] := 0.84130287;
      W_o[8,39] := -0.17293605;
      W_o[9,0] := -0.23097152;
      W_o[9,1] := -0.15871769;
      W_o[9,2] := 0.19358408;
      W_o[9,3] := -0.07425319;
      W_o[9,4] := -0.07420044;
      W_o[9,5] := -0.02661255;
      W_o[9,6] := 0.01253666;
      W_o[9,7] := 0.10329421;
      W_o[9,8] := -0.56111175;
      W_o[9,9] := -0.00908910;
      W_o[9,10] := 0.05690090;
      W_o[9,11] := -0.08010776;
      W_o[9,12] := -0.30403617;
      W_o[9,13] := 0.18955500;
      W_o[9,14] := 0.13771547;
      W_o[9,15] := -0.01777378;
      W_o[9,16] := -0.24138446;
      W_o[9,17] := -0.35579425;
      W_o[9,18] := -0.08040234;
      W_o[9,19] := -0.13508585;
      W_o[9,20] := -0.02945085;
      W_o[9,21] := 0.03336230;
      W_o[9,22] := -0.12277806;
      W_o[9,23] := -0.04557683;
      W_o[9,24] := -0.04875191;
      W_o[9,25] := -0.41637805;
      W_o[9,26] := -0.01602186;
      W_o[9,27] := 0.07369323;
      W_o[9,28] := 0.10504878;
      W_o[9,29] := 0.14198847;
      W_o[9,30] := 0.12163979;
      W_o[9,31] := -0.06927035;
      W_o[9,32] := 0.27943438;
      W_o[9,33] := 0.52821499;
      W_o[9,34] := -0.42556605;
      W_o[9,35] := -0.08720541;
      W_o[9,36] := -0.03627931;
      W_o[9,37] := -0.44218603;
      W_o[9,38] := 0.03999072;
      W_o[9,39] := 0.00299911;
      W_o[10,0] := -0.04975344;
      W_o[10,1] := -0.05351494;
      W_o[10,2] := -0.38371047;
      W_o[10,3] := -0.18595266;
      W_o[10,4] := 0.61007762;
      W_o[10,5] := 0.26893875;
      W_o[10,6] := 0.48405737;
      W_o[10,7] := 0.22436641;
      W_o[10,8] := 0.19901817;
      W_o[10,9] := -0.22706722;
      W_o[10,10] := -0.10738972;
      W_o[10,11] := -0.54268700;
      W_o[10,12] := 0.17331728;
      W_o[10,13] := 0.00065102;
      W_o[10,14] := 0.02936948;
      W_o[10,15] := -0.08635025;
      W_o[10,16] := -0.16275202;
      W_o[10,17] := 0.12818769;
      W_o[10,18] := -0.40466881;
      W_o[10,19] := 0.01480665;
      W_o[10,20] := -0.10567395;
      W_o[10,21] := -0.37431306;
      W_o[10,22] := -0.15547411;
      W_o[10,23] := -0.28764358;
      W_o[10,24] := 0.09085161;
      W_o[10,25] := 0.11554771;
      W_o[10,26] := -0.10251199;
      W_o[10,27] := 0.49218032;
      W_o[10,28] := -0.44367763;
      W_o[10,29] := 0.61115736;
      W_o[10,30] := 0.09082448;
      W_o[10,31] := -0.17321259;
      W_o[10,32] := -0.02935122;
      W_o[10,33] := -0.11259301;
      W_o[10,34] := 0.10632857;
      W_o[10,35] := -0.03293566;
      W_o[10,36] := -0.04883565;
      W_o[10,37] := -0.02677902;
      W_o[10,38] := 1.76672316;
      W_o[10,39] := 0.33624750;
      W_o[11,0] := 0.01394278;
      W_o[11,1] := 0.06421855;
      W_o[11,2] := -0.03070414;
      W_o[11,3] := -0.01582862;
      W_o[11,4] := 0.18139800;
      W_o[11,5] := 0.01746111;
      W_o[11,6] := -0.08357982;
      W_o[11,7] := 0.29224193;
      W_o[11,8] := -0.48481557;
      W_o[11,9] := 0.13723494;
      W_o[11,10] := -0.06989022;
      W_o[11,11] := 0.05515242;
      W_o[11,12] := 0.54017520;
      W_o[11,13] := -0.53452188;
      W_o[11,14] := -0.24097805;
      W_o[11,15] := 0.19763122;
      W_o[11,16] := 0.08363523;
      W_o[11,17] := 0.08858116;
      W_o[11,18] := -0.64370853;
      W_o[11,19] := -0.06206464;
      W_o[11,20] := -0.36461070;
      W_o[11,21] := -0.21325266;
      W_o[11,22] := -0.32683265;
      W_o[11,23] := -0.30821675;
      W_o[11,24] := -0.28392822;
      W_o[11,25] := -0.12898649;
      W_o[11,26] := 0.05272817;
      W_o[11,27] := 0.48492938;
      W_o[11,28] := -0.20675467;
      W_o[11,29] := 0.07431351;
      W_o[11,30] := -0.37345022;
      W_o[11,31] := 0.12173636;
      W_o[11,32] := -0.04922697;
      W_o[11,33] := -0.12817353;
      W_o[11,34] := -0.09397820;
      W_o[11,35] := 0.16107689;
      W_o[11,36] := -0.12483561;
      W_o[11,37] := 0.43916070;
      W_o[11,38] := -0.01915846;
      W_o[11,39] := 0.11393341;
      W_o[12,0] := 0.65769601;
      W_o[12,1] := 0.61452502;
      W_o[12,2] := 0.35834756;
      W_o[12,3] := -0.28856269;
      W_o[12,4] := -0.27414569;
      W_o[12,5] := -0.04396406;
      W_o[12,6] := -0.18361871;
      W_o[12,7] := -0.69043237;
      W_o[12,8] := 0.87575340;
      W_o[12,9] := -0.17673455;
      W_o[12,10] := -0.25065345;
      W_o[12,11] := -0.45248187;
      W_o[12,12] := -0.43163869;
      W_o[12,13] := 0.30214012;
      W_o[12,14] := 0.06767979;
      W_o[12,15] := -0.18445995;
      W_o[12,16] := 0.10103071;
      W_o[12,17] := 0.40537530;
      W_o[12,18] := 0.17058529;
      W_o[12,19] := 0.69663244;
      W_o[12,20] := -0.27960318;
      W_o[12,21] := 0.41710144;
      W_o[12,22] := 0.00595323;
      W_o[12,23] := 0.04762316;
      W_o[12,24] := -0.05134995;
      W_o[12,25] := 0.00458492;
      W_o[12,26] := -0.11405814;
      W_o[12,27] := -0.00941458;
      W_o[12,28] := 0.37036830;
      W_o[12,29] := 0.33941841;
      W_o[12,30] := -0.18241553;
      W_o[12,31] := 0.01994393;
      W_o[12,32] := -0.02669859;
      W_o[12,33] := 0.25948024;
      W_o[12,34] := 0.02076828;
      W_o[12,35] := -0.19220017;
      W_o[12,36] := -0.00991878;
      W_o[12,37] := 0.02291115;
      W_o[12,38] := 0.16625834;
      W_o[12,39] := -0.22731686;
      W_o[13,0] := -0.15924910;
      W_o[13,1] := -0.47062671;
      W_o[13,2] := 0.07512743;
      W_o[13,3] := -0.14161655;
      W_o[13,4] := 0.30482900;
      W_o[13,5] := -0.31820074;
      W_o[13,6] := 0.42128560;
      W_o[13,7] := 0.04020222;
      W_o[13,8] := 0.64258534;
      W_o[13,9] := 0.31215358;
      W_o[13,10] := -0.37166351;
      W_o[13,11] := -0.12368796;
      W_o[13,12] := -0.02779209;
      W_o[13,13] := -0.86361456;
      W_o[13,14] := 0.01958641;
      W_o[13,15] := 0.05256082;
      W_o[13,16] := -0.07068108;
      W_o[13,17] := 0.04328666;
      W_o[13,18] := 0.34329355;
      W_o[13,19] := -0.57730550;
      W_o[13,20] := -0.19776343;
      W_o[13,21] := -0.17221977;
      W_o[13,22] := 0.09852456;
      W_o[13,23] := -1.00299084;
      W_o[13,24] := 2.34005952;
      W_o[13,25] := 1.83858848;
      W_o[13,26] := -0.86023897;
      W_o[13,27] := 0.10414210;
      W_o[13,28] := -0.38447699;
      W_o[13,29] := 0.01457757;
      W_o[13,30] := 0.18932407;
      W_o[13,31] := 0.56862438;
      W_o[13,32] := 0.08322045;
      W_o[13,33] := -0.18533768;
      W_o[13,34] := 1.10703778;
      W_o[13,35] := -0.28043205;
      W_o[13,36] := -0.30521935;
      W_o[13,37] := -0.34443730;
      W_o[13,38] := -0.01801103;
      W_o[13,39] := -0.13203925;
      W_o[14,0] := -0.02214651;
      W_o[14,1] := 0.41877946;
      W_o[14,2] := -0.21624404;
      W_o[14,3] := 0.59027672;
      W_o[14,4] := 0.29192978;
      W_o[14,5] := 0.70612335;
      W_o[14,6] := 0.69886094;
      W_o[14,7] := 0.43926716;
      W_o[14,8] := -0.70507145;
      W_o[14,9] := 0.46977445;
      W_o[14,10] := 0.50927150;
      W_o[14,11] := -0.12555990;
      W_o[14,12] := -0.03891997;
      W_o[14,13] := 0.45297027;
      W_o[14,14] := 0.10233755;
      W_o[14,15] := -0.29167077;
      W_o[14,16] := -0.12342054;
      W_o[14,17] := 0.00189050;
      W_o[14,18] := 0.16054912;
      W_o[14,19] := -0.00484559;
      W_o[14,20] := -0.36701992;
      W_o[14,21] := -0.05176546;
      W_o[14,22] := 0.00353710;
      W_o[14,23] := -0.00093972;
      W_o[14,24] := 0.32338837;
      W_o[14,25] := 0.28439587;
      W_o[14,26] := -0.08737835;
      W_o[14,27] := -0.04817959;
      W_o[14,28] := 0.18409094;
      W_o[14,29] := -0.03510422;
      W_o[14,30] := -0.01086587;
      W_o[14,31] := 0.02054300;
      W_o[14,32] := -0.07345553;
      W_o[14,33] := -0.21690357;
      W_o[14,34] := -0.28374419;
      W_o[14,35] := 0.02088533;
      W_o[14,36] := 0.07017583;
      W_o[14,37] := -0.12823847;
      W_o[14,38] := 0.25906608;
      W_o[14,39] := -0.18490438;
      W_o[15,0] := 0.00456393;
      W_o[15,1] := 0.20027003;
      W_o[15,2] := -0.10480183;
      W_o[15,3] := 0.31756738;
      W_o[15,4] := -0.10564005;
      W_o[15,5] := 0.02531332;
      W_o[15,6] := 0.32546297;
      W_o[15,7] := -0.03057292;
      W_o[15,8] := -0.09481000;
      W_o[15,9] := 0.00536214;
      W_o[15,10] := 0.12456731;
      W_o[15,11] := 0.08706652;
      W_o[15,12] := 0.19711065;
      W_o[15,13] := -0.11705462;
      W_o[15,14] := -0.00124244;
      W_o[15,15] := -0.66989708;
      W_o[15,16] := 0.18187341;
      W_o[15,17] := 0.00445009;
      W_o[15,18] := 2.26799989;
      W_o[15,19] := -0.33114424;
      W_o[15,20] := 0.08577366;
      W_o[15,21] := 0.26837903;
      W_o[15,22] := 0.10760636;
      W_o[15,23] := -0.22246659;
      W_o[15,24] := -0.21526244;
      W_o[15,25] := 0.00395280;
      W_o[15,26] := 0.03160953;
      W_o[15,27] := -0.39023194;
      W_o[15,28] := 0.21006531;
      W_o[15,29] := 0.34472552;
      W_o[15,30] := 0.31186867;
      W_o[15,31] := 0.00415714;
      W_o[15,32] := 0.23063444;
      W_o[15,33] := 0.19425058;
      W_o[15,34] := 0.27053815;
      W_o[15,35] := 0.17631577;
      W_o[15,36] := 0.04783322;
      W_o[15,37] := 0.08611892;
      W_o[15,38] := 0.38180444;
      W_o[15,39] := -0.20466073;
      W_o[16,0] := -0.15114191;
      W_o[16,1] := 0.00804333;
      W_o[16,2] := 0.06051351;
      W_o[16,3] := 0.28815919;
      W_o[16,4] := 0.18742214;
      W_o[16,5] := -0.11313698;
      W_o[16,6] := -0.13429113;
      W_o[16,7] := -0.23928368;
      W_o[16,8] := -0.29211384;
      W_o[16,9] := 0.30963427;
      W_o[16,10] := 0.01700113;
      W_o[16,11] := -0.16528781;
      W_o[16,12] := -0.08125683;
      W_o[16,13] := -0.04685068;
      W_o[16,14] := 0.82725412;
      W_o[16,15] := -0.02709327;
      W_o[16,16] := -0.03765779;
      W_o[16,17] := -0.54237044;
      W_o[16,18] := -0.01633970;
      W_o[16,19] := 1.70895028;
      W_o[16,20] := -0.21961294;
      W_o[16,21] := -0.07729631;
      W_o[16,22] := -0.04895397;
      W_o[16,23] := 0.01796570;
      W_o[16,24] := 0.10057043;
      W_o[16,25] := 0.08332445;
      W_o[16,26] := -0.01614249;
      W_o[16,27] := -0.05278811;
      W_o[16,28] := -0.12061049;
      W_o[16,29] := 0.09612570;
      W_o[16,30] := -0.27439341;
      W_o[16,31] := 0.02516360;
      W_o[16,32] := -0.17176309;
      W_o[16,33] := -0.05478594;
      W_o[16,34] := -0.00976936;
      W_o[16,35] := -0.15284751;
      W_o[16,36] := 0.00708155;
      W_o[16,37] := -0.10585996;
      W_o[16,38] := 0.09140552;
      W_o[16,39] := -0.26013094;
      W_o[17,0] := 0.08286103;
      W_o[17,1] := 0.03750033;
      W_o[17,2] := -0.10766149;
      W_o[17,3] := 0.61591530;
      W_o[17,4] := -0.14656810;
      W_o[17,5] := -0.02154700;
      W_o[17,6] := -0.08073130;
      W_o[17,7] := -0.05106850;
      W_o[17,8] := 0.01058245;
      W_o[17,9] := -0.36430576;
      W_o[17,10] := -0.23940334;
      W_o[17,11] := -0.51427031;
      W_o[17,12] := 0.67015946;
      W_o[17,13] := -0.10680982;
      W_o[17,14] := -0.02610255;
      W_o[17,15] := -0.15557665;
      W_o[17,16] := 0.10917784;
      W_o[17,17] := -0.02499565;
      W_o[17,18] := -0.03614269;
      W_o[17,19] := -0.47785047;
      W_o[17,20] := -0.18451281;
      W_o[17,21] := 0.10915274;
      W_o[17,22] := -0.36744645;
      W_o[17,23] := -0.10975158;
      W_o[17,24] := 0.21045783;
      W_o[17,25] := 0.09130947;
      W_o[17,26] := 0.01529007;
      W_o[17,27] := -0.18475625;
      W_o[17,28] := 0.08889312;
      W_o[17,29] := 0.05933971;
      W_o[17,30] := -0.31048802;
      W_o[17,31] := -0.03528069;
      W_o[17,32] := -0.20060484;
      W_o[17,33] := 0.33930284;
      W_o[17,34] := 0.22307321;
      W_o[17,35] := -0.12793279;
      W_o[17,36] := 0.03892962;
      W_o[17,37] := -0.39412618;
      W_o[17,38] := 1.05452859;
      W_o[17,39] := 0.05015264;
      W_o[18,0] := 0.61441380;
      W_o[18,1] := -0.00581962;
      W_o[18,2] := 0.01838240;
      W_o[18,3] := 0.17021340;
      W_o[18,4] := -0.14046310;
      W_o[18,5] := -0.03963570;
      W_o[18,6] := -0.16133307;
      W_o[18,7] := -0.08786807;
      W_o[18,8] := 0.66064078;
      W_o[18,9] := -0.50882161;
      W_o[18,10] := 0.05472949;
      W_o[18,11] := -0.40465507;
      W_o[18,12] := -0.16453871;
      W_o[18,13] := -0.07766686;
      W_o[18,14] := 0.03071279;
      W_o[18,15] := -0.08571735;
      W_o[18,16] := -0.11585758;
      W_o[18,17] := 0.10421877;
      W_o[18,18] := -0.30685908;
      W_o[18,19] := -0.72102994;
      W_o[18,20] := -0.39853510;
      W_o[18,21] := -0.47263488;
      W_o[18,22] := -0.65301901;
      W_o[18,23] := 0.04909870;
      W_o[18,24] := -0.26901412;
      W_o[18,25] := -0.43715164;
      W_o[18,26] := -0.33605048;
      W_o[18,27] := 0.12228665;
      W_o[18,28] := 0.31939563;
      W_o[18,29] := 0.21070679;
      W_o[18,30] := -0.58367223;
      W_o[18,31] := 0.44466385;
      W_o[18,32] := 0.11434247;
      W_o[18,33] := 0.13122903;
      W_o[18,34] := -0.08403879;
      W_o[18,35] := 0.23515210;
      W_o[18,36] := 0.09416876;
      W_o[18,37] := 0.43245336;
      W_o[18,38] := 0.42059562;
      W_o[18,39] := -0.27610445;
      W_o[19,0] := -0.34880528;
      W_o[19,1] := -0.11340433;
      W_o[19,2] := 0.00313819;
      W_o[19,3] := 0.61080855;
      W_o[19,4] := 0.09961273;
      W_o[19,5] := 0.15991150;
      W_o[19,6] := -0.17713304;
      W_o[19,7] := 0.17079115;
      W_o[19,8] := 0.10543557;
      W_o[19,9] := -0.38165331;
      W_o[19,10] := 0.08110224;
      W_o[19,11] := 0.12665251;
      W_o[19,12] := 0.76474392;
      W_o[19,13] := -0.97162247;
      W_o[19,14] := -0.15689284;
      W_o[19,15] := -0.15970281;
      W_o[19,16] := 0.26374424;
      W_o[19,17] := -0.16025481;
      W_o[19,18] := -0.48080701;
      W_o[19,19] := -0.51185387;
      W_o[19,20] := -0.10991344;
      W_o[19,21] := -0.05593008;
      W_o[19,22] := -0.15545925;
      W_o[19,23] := -0.43545204;
      W_o[19,24] := 1.16323590;
      W_o[19,25] := 1.17089522;
      W_o[19,26] := 0.07496043;
      W_o[19,27] := 0.46996966;
      W_o[19,28] := 0.14273608;
      W_o[19,29] := -0.10301508;
      W_o[19,30] := -0.17604618;
      W_o[19,31] := -0.18035652;
      W_o[19,32] := -0.17284030;
      W_o[19,33] := -0.21061423;
      W_o[19,34] := -0.48001161;
      W_o[19,35] := 0.15144287;
      W_o[19,36] := -0.10487883;
      W_o[19,37] := 0.21051478;
      W_o[19,38] := -0.03737800;
      W_o[19,39] := 0.22113863;
      W_o[20,0] := -0.09744378;
      W_o[20,1] := -0.01674240;
      W_o[20,2] := 0.01145337;
      W_o[20,3] := -0.16928835;
      W_o[20,4] := -0.08487850;
      W_o[20,5] := 0.16698468;
      W_o[20,6] := -0.63689768;
      W_o[20,7] := 0.33002836;
      W_o[20,8] := -0.74119657;
      W_o[20,9] := 0.52214622;
      W_o[20,10] := -0.66047299;
      W_o[20,11] := -0.43090153;
      W_o[20,12] := -0.27590305;
      W_o[20,13] := 0.15499099;
      W_o[20,14] := 0.11995452;
      W_o[20,15] := -0.02210920;
      W_o[20,16] := 0.06650748;
      W_o[20,17] := 0.00387770;
      W_o[20,18] := 0.48246086;
      W_o[20,19] := -0.01958447;
      W_o[20,20] := 0.12180612;
      W_o[20,21] := 0.24685419;
      W_o[20,22] := -0.13427232;
      W_o[20,23] := 0.06217969;
      W_o[20,24] := 1.25715184;
      W_o[20,25] := 0.77083719;
      W_o[20,26] := -0.31976116;
      W_o[20,27] := 0.18783310;
      W_o[20,28] := -0.05193661;
      W_o[20,29] := 0.09904788;
      W_o[20,30] := -0.12382533;
      W_o[20,31] := 0.04432494;
      W_o[20,32] := -0.07709737;
      W_o[20,33] := 0.00720727;
      W_o[20,34] := 0.14193270;
      W_o[20,35] := -0.18251143;
      W_o[20,36] := -0.00754279;
      W_o[20,37] := -0.16062810;
      W_o[20,38] := -0.09272868;
      W_o[20,39] := -0.15935695;
      W_o[21,0] := -0.22163987;
      W_o[21,1] := -0.07309268;
      W_o[21,2] := -0.03787788;
      W_o[21,3] := 0.28699502;
      W_o[21,4] := 0.18230651;
      W_o[21,5] := -0.30771858;
      W_o[21,6] := -0.03588717;
      W_o[21,7] := 0.20533676;
      W_o[21,8] := -0.08486333;
      W_o[21,9] := -0.01344010;
      W_o[21,10] := -0.52408534;
      W_o[21,11] := 0.02502864;
      W_o[21,12] := -0.83751518;
      W_o[21,13] := -0.03175629;
      W_o[21,14] := 0.21095377;
      W_o[21,15] := -0.84907478;
      W_o[21,16] := 0.00443229;
      W_o[21,17] := 0.24032350;
      W_o[21,18] := 0.20381300;
      W_o[21,19] := -0.53694773;
      W_o[21,20] := -0.09315480;
      W_o[21,21] := -0.33405665;
      W_o[21,22] := 0.05652494;
      W_o[21,23] := 0.36037019;
      W_o[21,24] := 0.20759679;
      W_o[21,25] := 0.06819481;
      W_o[21,26] := 0.13676454;
      W_o[21,27] := 0.64053833;
      W_o[21,28] := 0.11439332;
      W_o[21,29] := -0.37118480;
      W_o[21,30] := -0.00156529;
      W_o[21,31] := -0.07878110;
      W_o[21,32] := -0.21185711;
      W_o[21,33] := -0.09498084;
      W_o[21,34] := -0.12056343;
      W_o[21,35] := -0.28038767;
      W_o[21,36] := 0.00132361;
      W_o[21,37] := -0.09131619;
      W_o[21,38] := -0.27713600;
      W_o[21,39] := -0.28789780;
      W_o[22,0] := -0.15200722;
      W_o[22,1] := 0.80616361;
      W_o[22,2] := 0.09922904;
      W_o[22,3] := -0.20402044;
      W_o[22,4] := 0.10210901;
      W_o[22,5] := 0.09848336;
      W_o[22,6] := -0.19488986;
      W_o[22,7] := 0.07671145;
      W_o[22,8] := -0.20990044;
      W_o[22,9] := 0.08224703;
      W_o[22,10] := 0.20208466;
      W_o[22,11] := 0.02182630;
      W_o[22,12] := -0.17363830;
      W_o[22,13] := 0.25162092;
      W_o[22,14] := -0.24746750;
      W_o[22,15] := -0.12957299;
      W_o[22,16] := -0.00627271;
      W_o[22,17] := 0.03615937;
      W_o[22,18] := 0.33972406;
      W_o[22,19] := 0.11538468;
      W_o[22,20] := 0.04234114;
      W_o[22,21] := 0.47518721;
      W_o[22,22] := 0.41847426;
      W_o[22,23] := -0.35500267;
      W_o[22,24] := 1.08033085;
      W_o[22,25] := 1.00722659;
      W_o[22,26] := -0.28602570;
      W_o[22,27] := -0.06139164;
      W_o[22,28] := 0.05762752;
      W_o[22,29] := 0.09372402;
      W_o[22,30] := 0.42476979;
      W_o[22,31] := 0.13689539;
      W_o[22,32] := 0.25176939;
      W_o[22,33] := 0.23804808;
      W_o[22,34] := 0.38350585;
      W_o[22,35] := 0.14343651;
      W_o[22,36] := -0.01567702;
      W_o[22,37] := 0.41862074;
      W_o[22,38] := -0.02235131;
      W_o[22,39] := 1.10857010;
      W_o[23,0] := 0.29647908;
      W_o[23,1] := -0.09007457;
      W_o[23,2] := -0.51309329;
      W_o[23,3] := -0.32924581;
      W_o[23,4] := -0.16417709;
      W_o[23,5] := 0.05021456;
      W_o[23,6] := 0.09369662;
      W_o[23,7] := -0.09293582;
      W_o[23,8] := -0.06115354;
      W_o[23,9] := 0.47681352;
      W_o[23,10] := 0.11118036;
      W_o[23,11] := -0.36791933;
      W_o[23,12] := -0.64249408;
      W_o[23,13] := 0.16806115;
      W_o[23,14] := 0.05251247;
      W_o[23,15] := -0.44162959;
      W_o[23,16] := -0.03784051;
      W_o[23,17] := 0.01734663;
      W_o[23,18] := -0.05495093;
      W_o[23,19] := -0.09302599;
      W_o[23,20] := 0.21550827;
      W_o[23,21] := 0.02342126;
      W_o[23,22] := -0.65106291;
      W_o[23,23] := -0.16059713;
      W_o[23,24] := 0.74768978;
      W_o[23,25] := 0.77801579;
      W_o[23,26] := -0.13329148;
      W_o[23,27] := -0.01115259;
      W_o[23,28] := 0.20939310;
      W_o[23,29] := -0.14855206;
      W_o[23,30] := -0.59163791;
      W_o[23,31] := -0.10205384;
      W_o[23,32] := -0.17358899;
      W_o[23,33] := 0.19429116;
      W_o[23,34] := -0.44206089;
      W_o[23,35] := -0.13230647;
      W_o[23,36] := -0.00379825;
      W_o[23,37] := -0.31613481;
      W_o[23,38] := -0.03437910;
      W_o[23,39] := 0.69593823;
      W_o[24,0] := 0.18129924;
      W_o[24,1] := 0.63154942;
      W_o[24,2] := -0.01074047;
      W_o[24,3] := 0.30104062;
      W_o[24,4] := 0.07274275;
      W_o[24,5] := -0.20634146;
      W_o[24,6] := 0.07617958;
      W_o[24,7] := -0.09617994;
      W_o[24,8] := 0.02491149;
      W_o[24,9] := -0.01619528;
      W_o[24,10] := 0.74655634;
      W_o[24,11] := -0.32350552;
      W_o[24,12] := -0.18770587;
      W_o[24,13] := -0.17258902;
      W_o[24,14] := -0.13972870;
      W_o[24,15] := -0.77128297;
      W_o[24,16] := 0.14157821;
      W_o[24,17] := -0.05731640;
      W_o[24,18] := 0.19687349;
      W_o[24,19] := -0.30524209;
      W_o[24,20] := -0.24232426;
      W_o[24,21] := 0.12608968;
      W_o[24,22] := 0.01551487;
      W_o[24,23] := -0.41677731;
      W_o[24,24] := 0.93884945;
      W_o[24,25] := 0.78144521;
      W_o[24,26] := -0.38716099;
      W_o[24,27] := -0.01172645;
      W_o[24,28] := 0.00427037;
      W_o[24,29] := -0.10702599;
      W_o[24,30] := -0.06169849;
      W_o[24,31] := -0.04865468;
      W_o[24,32] := -0.21641125;
      W_o[24,33] := -0.27539209;
      W_o[24,34] := 0.78715312;
      W_o[24,35] := -0.14164442;
      W_o[24,36] := -0.17446344;
      W_o[24,37] := 0.05613173;
      W_o[24,38] := 0.25165775;
      W_o[24,39] := 0.32816496;
      W_o[25,0] := -0.09599993;
      W_o[25,1] := -0.25011954;
      W_o[25,2] := -0.03694122;
      W_o[25,3] := -0.62371397;
      W_o[25,4] := 0.23611289;
      W_o[25,5] := 0.28173044;
      W_o[25,6] := -0.30132398;
      W_o[25,7] := 0.39865136;
      W_o[25,8] := -0.09741599;
      W_o[25,9] := -0.25187540;
      W_o[25,10] := 0.27679303;
      W_o[25,11] := -0.27845952;
      W_o[25,12] := -0.06051615;
      W_o[25,13] := -0.11906760;
      W_o[25,14] := -0.13467777;
      W_o[25,15] := -0.15183683;
      W_o[25,16] := 0.01077802;
      W_o[25,17] := -0.15232092;
      W_o[25,18] := 0.31490743;
      W_o[25,19] := 0.06639913;
      W_o[25,20] := -0.68352765;
      W_o[25,21] := 0.32349935;
      W_o[25,22] := -0.02829045;
      W_o[25,23] := 0.09799626;
      W_o[25,24] := -0.41351509;
      W_o[25,25] := -0.43447980;
      W_o[25,26] := 0.18629681;
      W_o[25,27] := 0.59058458;
      W_o[25,28] := -0.06618728;
      W_o[25,29] := 1.18627656;
      W_o[25,30] := -0.04305683;
      W_o[25,31] := -0.16967137;
      W_o[25,32] := 0.27466226;
      W_o[25,33] := 0.06906415;
      W_o[25,34] := -0.33705801;
      W_o[25,35] := -0.17390864;
      W_o[25,36] := -0.13643852;
      W_o[25,37] := 0.15441231;
      W_o[25,38] := -0.15764047;
      W_o[25,39] := 0.03892670;
      W_o[26,0] := 0.14575106;
      W_o[26,1] := 0.63006645;
      W_o[26,2] := -0.19157562;
      W_o[26,3] := -0.00748385;
      W_o[26,4] := 0.01923200;
      W_o[26,5] := 0.09620106;
      W_o[26,6] := 0.13181686;
      W_o[26,7] := 0.19512504;
      W_o[26,8] := 0.19447267;
      W_o[26,9] := 0.07103106;
      W_o[26,10] := -0.25106451;
      W_o[26,11] := 0.07562301;
      W_o[26,12] := 0.16949712;
      W_o[26,13] := 0.77973145;
      W_o[26,14] := -0.00400880;
      W_o[26,15] := -0.30748934;
      W_o[26,16] := -0.04597035;
      W_o[26,17] := -0.11540623;
      W_o[26,18] := 0.61029083;
      W_o[26,19] := -0.13811298;
      W_o[26,20] := -0.44542348;
      W_o[26,21] := 0.55551034;
      W_o[26,22] := -0.07641070;
      W_o[26,23] := 0.06676203;
      W_o[26,24] := 0.00876335;
      W_o[26,25] := -0.08375374;
      W_o[26,26] := -0.46028519;
      W_o[26,27] := 0.41610366;
      W_o[26,28] := -0.06305913;
      W_o[26,29] := 0.01283880;
      W_o[26,30] := 0.00893430;
      W_o[26,31] := 0.11318304;
      W_o[26,32] := -0.00202851;
      W_o[26,33] := 0.06692720;
      W_o[26,34] := 0.08405498;
      W_o[26,35] := -0.13670896;
      W_o[26,36] := 0.01352034;
      W_o[26,37] := -0.13026740;
      W_o[26,38] := 0.65490270;
      W_o[26,39] := -0.08570544;
      W_o[27,0] := -0.11447388;
      W_o[27,1] := -0.42843413;
      W_o[27,2] := -0.04269759;
      W_o[27,3] := -0.40117773;
      W_o[27,4] := -0.24858794;
      W_o[27,5] := -0.04377360;
      W_o[27,6] := -0.39127943;
      W_o[27,7] := -0.51688462;
      W_o[27,8] := 0.07314450;
      W_o[27,9] := -0.21077925;
      W_o[27,10] := -0.22803664;
      W_o[27,11] := 0.08533891;
      W_o[27,12] := -0.18755989;
      W_o[27,13] := 0.24690123;
      W_o[27,14] := 0.02400121;
      W_o[27,15] := 0.02479623;
      W_o[27,16] := 0.04027365;
      W_o[27,17] := -0.00776743;
      W_o[27,18] := 0.75450927;
      W_o[27,19] := -0.06382228;
      W_o[27,20] := -0.23799492;
      W_o[27,21] := -0.18352440;
      W_o[27,22] := -0.37799615;
      W_o[27,23] := -0.77834731;
      W_o[27,24] := 0.79094517;
      W_o[27,25] := 0.37767863;
      W_o[27,26] := 0.45343819;
      W_o[27,27] := 0.27995503;
      W_o[27,28] := 0.04575095;
      W_o[27,29] := -0.40213665;
      W_o[27,30] := -0.61576760;
      W_o[27,31] := -0.01314038;
      W_o[27,32] := -0.19220178;
      W_o[27,33] := -0.18640390;
      W_o[27,34] := -1.05954719;
      W_o[27,35] := -0.31399265;
      W_o[27,36] := -0.08189996;
      W_o[27,37] := -0.26056018;
      W_o[27,38] := -0.15719463;
      W_o[27,39] := -0.03270736;
      W_o[28,0] := 0.28491798;
      W_o[28,1] := 0.23311718;
      W_o[28,2] := 0.09096937;
      W_o[28,3] := -0.38070893;
      W_o[28,4] := 0.33497691;
      W_o[28,5] := 0.02360616;
      W_o[28,6] := -0.40364549;
      W_o[28,7] := 0.52994388;
      W_o[28,8] := 0.18476413;
      W_o[28,9] := -0.41934469;
      W_o[28,10] := 0.09743979;
      W_o[28,11] := -0.06271173;
      W_o[28,12] := -0.33278829;
      W_o[28,13] := 0.09721936;
      W_o[28,14] := 0.05886953;
      W_o[28,15] := -0.02753331;
      W_o[28,16] := -0.28607798;
      W_o[28,17] := -0.10859327;
      W_o[28,18] := -0.19896559;
      W_o[28,19] := -0.33864468;
      W_o[28,20] := -0.11514115;
      W_o[28,21] := 0.22684307;
      W_o[28,22] := -0.07266788;
      W_o[28,23] := -0.00887611;
      W_o[28,24] := -0.03110049;
      W_o[28,25] := 0.42423946;
      W_o[28,26] := 0.16166633;
      W_o[28,27] := 0.46223441;
      W_o[28,28] := 0.15797591;
      W_o[28,29] := 0.18892875;
      W_o[28,30] := -0.06017169;
      W_o[28,31] := 0.01324773;
      W_o[28,32] := 0.10118480;
      W_o[28,33] := 0.08109213;
      W_o[28,34] := -0.05838856;
      W_o[28,35] := 0.27322558;
      W_o[28,36] := -0.01824474;
      W_o[28,37] := 0.21420285;
      W_o[28,38] := 0.17817383;
      W_o[28,39] := 0.09010561;
      W_o[29,0] := 0.07731791;
      W_o[29,1] := -0.09667790;
      W_o[29,2] := -0.07639322;
      W_o[29,3] := -0.05219271;
      W_o[29,4] := 0.05173031;
      W_o[29,5] := 0.20557168;
      W_o[29,6] := -0.08309768;
      W_o[29,7] := -0.11951208;
      W_o[29,8] := 0.04824584;
      W_o[29,9] := 0.00393840;
      W_o[29,10] := -0.01744876;
      W_o[29,11] := -0.02404173;
      W_o[29,12] := 0.09710021;
      W_o[29,13] := -0.01241371;
      W_o[29,14] := -0.01065864;
      W_o[29,15] := -0.04493345;
      W_o[29,16] := -0.00543620;
      W_o[29,17] := 0.01306327;
      W_o[29,18] := 0.01685135;
      W_o[29,19] := -0.04317724;
      W_o[29,20] := -0.06109453;
      W_o[29,21] := -0.25755301;
      W_o[29,22] := -0.10231650;
      W_o[29,23] := 0.02879286;
      W_o[29,24] := -0.56473893;
      W_o[29,25] := -0.54539061;
      W_o[29,26] := -0.17247662;
      W_o[29,27] := 0.24084187;
      W_o[29,28] := -0.10003161;
      W_o[29,29] := -0.41303715;
      W_o[29,30] := -0.10672592;
      W_o[29,31] := -0.05027681;
      W_o[29,32] := -0.14264677;
      W_o[29,33] := -0.11566567;
      W_o[29,34] := -0.53422034;
      W_o[29,35] := -0.05037379;
      W_o[29,36] := -0.01575625;
      W_o[29,37] := -0.11289191;
      W_o[29,38] := 0.00716874;
      W_o[29,39] := 1.32865441;
      W_o[30,0] := -0.17489706;
      W_o[30,1] := -0.04965573;
      W_o[30,2] := 0.10585558;
      W_o[30,3] := 0.77944791;
      W_o[30,4] := -0.04518570;
      W_o[30,5] := -0.18553282;
      W_o[30,6] := 0.08056828;
      W_o[30,7] := -0.20592566;
      W_o[30,8] := -0.06633148;
      W_o[30,9] := -0.53728795;
      W_o[30,10] := 0.04003848;
      W_o[30,11] := -0.28942955;
      W_o[30,12] := -0.63946211;
      W_o[30,13] := 0.26434416;
      W_o[30,14] := -0.06438407;
      W_o[30,15] := -0.94219506;
      W_o[30,16] := -0.09090893;
      W_o[30,17] := -0.24020159;
      W_o[30,18] := 1.13913250;
      W_o[30,19] := 0.09926897;
      W_o[30,20] := 0.02266491;
      W_o[30,21] := -0.07792678;
      W_o[30,22] := -0.01553794;
      W_o[30,23] := -0.10481242;
      W_o[30,24] := -0.15663289;
      W_o[30,25] := -0.12417895;
      W_o[30,26] := -0.16360331;
      W_o[30,27] := 0.09446005;
      W_o[30,28] := 0.13794288;
      W_o[30,29] := -0.17225608;
      W_o[30,30] := 0.04900527;
      W_o[30,31] := 0.39925125;
      W_o[30,32] := -0.08859237;
      W_o[30,33] := -0.06575945;
      W_o[30,34] := -0.20326042;
      W_o[30,35] := -0.02266855;
      W_o[30,36] := 0.03377234;
      W_o[30,37] := -0.13112211;
      W_o[30,38] := -0.05310003;
      W_o[30,39] := 0.83231968;
      W_o[31,0] := 0.15999089;
      W_o[31,1] := -0.05416152;
      W_o[31,2] := -0.07443288;
      W_o[31,3] := -0.19782902;
      W_o[31,4] := 0.08784235;
      W_o[31,5] := 0.09198477;
      W_o[31,6] := -0.19657053;
      W_o[31,7] := -0.05733800;
      W_o[31,8] := 0.03709866;
      W_o[31,9] := 0.02747005;
      W_o[31,10] := -0.15585202;
      W_o[31,11] := -0.54856622;
      W_o[31,12] := -0.37941724;
      W_o[31,13] := 0.18906285;
      W_o[31,14] := 0.01572132;
      W_o[31,15] := -0.53865492;
      W_o[31,16] := -0.47697246;
      W_o[31,17] := 0.07002753;
      W_o[31,18] := 0.55318737;
      W_o[31,19] := -0.15192324;
      W_o[31,20] := -0.04416887;
      W_o[31,21] := -0.07441948;
      W_o[31,22] := -0.02111035;
      W_o[31,23] := -0.12010260;
      W_o[31,24] := 1.28149831;
      W_o[31,25] := 0.69010407;
      W_o[31,26] := -0.05445243;
      W_o[31,27] := 0.17313376;
      W_o[31,28] := -0.03698421;
      W_o[31,29] := 0.75948030;
      W_o[31,30] := 0.00256974;
      W_o[31,31] := 0.01054981;
      W_o[31,32] := 0.14877367;
      W_o[31,33] := 0.08370097;
      W_o[31,34] := 0.13622369;
      W_o[31,35] := 0.05027818;
      W_o[31,36] := -0.06672458;
      W_o[31,37] := 0.18186426;
      W_o[31,38] := 0.06507517;
      W_o[31,39] := -0.35338154;
      R_i[0,0] := 0.02777663;
      R_i[0,1] := -0.30641955;
      R_i[0,2] := 0.11692245;
      R_i[0,3] := 0.29124752;
      R_i[0,4] := 0.05408674;
      R_i[0,5] := -0.13721205;
      R_i[0,6] := 0.54630709;
      R_i[0,7] := -0.27012211;
      R_i[0,8] := 0.15503287;
      R_i[0,9] := 0.10762413;
      R_i[0,10] := 0.17625292;
      R_i[0,11] := -0.04361302;
      R_i[0,12] := -0.08274892;
      R_i[0,13] := -0.14828911;
      R_i[0,14] := -0.19601791;
      R_i[0,15] := 0.30961239;
      R_i[0,16] := -0.28616810;
      R_i[0,17] := 0.37507176;
      R_i[0,18] := -0.04757742;
      R_i[0,19] := -0.00805486;
      R_i[0,20] := -0.19719143;
      R_i[0,21] := -0.20838951;
      R_i[0,22] := 0.01867366;
      R_i[0,23] := 0.14011624;
      R_i[0,24] := -0.17484367;
      R_i[0,25] := -0.14716677;
      R_i[0,26] := 0.27535814;
      R_i[0,27] := -0.26792911;
      R_i[0,28] := 0.13091210;
      R_i[0,29] := -0.00004443;
      R_i[0,30] := -0.31875929;
      R_i[0,31] := -0.23393498;
      R_i[1,0] := 0.09890532;
      R_i[1,1] := -0.41096249;
      R_i[1,2] := 0.22243534;
      R_i[1,3] := 0.28512338;
      R_i[1,4] := 0.15052673;
      R_i[1,5] := 0.08439466;
      R_i[1,6] := 0.13953692;
      R_i[1,7] := -0.06284653;
      R_i[1,8] := -0.15906256;
      R_i[1,9] := -0.02961123;
      R_i[1,10] := -0.07504162;
      R_i[1,11] := -0.05802333;
      R_i[1,12] := -0.01100338;
      R_i[1,13] := 0.09784974;
      R_i[1,14] := 0.21630995;
      R_i[1,15] := 0.03157408;
      R_i[1,16] := -0.14952427;
      R_i[1,17] := 0.21040013;
      R_i[1,18] := 0.73434794;
      R_i[1,19] := -0.18868551;
      R_i[1,20] := -0.02286376;
      R_i[1,21] := -0.09064758;
      R_i[1,22] := -0.32558787;
      R_i[1,23] := 0.07301825;
      R_i[1,24] := -0.09908721;
      R_i[1,25] := -0.22047330;
      R_i[1,26] := 0.18392785;
      R_i[1,27] := 0.29104322;
      R_i[1,28] := 0.65344906;
      R_i[1,29] := -0.07514935;
      R_i[1,30] := -0.17124803;
      R_i[1,31] := -0.07562800;
      R_i[2,0] := -0.18058190;
      R_i[2,1] := -0.09578291;
      R_i[2,2] := 0.14311229;
      R_i[2,3] := -0.16814849;
      R_i[2,4] := 0.22336932;
      R_i[2,5] := 0.08362369;
      R_i[2,6] := -0.01463015;
      R_i[2,7] := 0.04053539;
      R_i[2,8] := -0.22425680;
      R_i[2,9] := 0.30432880;
      R_i[2,10] := -0.04152664;
      R_i[2,11] := -0.12698807;
      R_i[2,12] := 0.04107983;
      R_i[2,13] := -0.07066728;
      R_i[2,14] := -0.32119438;
      R_i[2,15] := 0.19552983;
      R_i[2,16] := -0.40282956;
      R_i[2,17] := 0.21768214;
      R_i[2,18] := 0.11086221;
      R_i[2,19] := 0.03130512;
      R_i[2,20] := 0.27946118;
      R_i[2,21] := 0.15343487;
      R_i[2,22] := -0.16819488;
      R_i[2,23] := 0.05245676;
      R_i[2,24] := -0.04345716;
      R_i[2,25] := -0.45481893;
      R_i[2,26] := 0.10744009;
      R_i[2,27] := -0.16157587;
      R_i[2,28] := -0.27564815;
      R_i[2,29] := 0.29775959;
      R_i[2,30] := -0.30921066;
      R_i[2,31] := -0.17098905;
      R_i[3,0] := 0.23412624;
      R_i[3,1] := -0.32581827;
      R_i[3,2] := -0.04527292;
      R_i[3,3] := 1.06161284;
      R_i[3,4] := -0.10460636;
      R_i[3,5] := -0.01773712;
      R_i[3,6] := 0.42387381;
      R_i[3,7] := -0.02749722;
      R_i[3,8] := -0.39747861;
      R_i[3,9] := 0.33761570;
      R_i[3,10] := 0.91908520;
      R_i[3,11] := -0.12909365;
      R_i[3,12] := 0.12688540;
      R_i[3,13] := -0.16723385;
      R_i[3,14] := -0.16277122;
      R_i[3,15] := -0.37805018;
      R_i[3,16] := -0.15600394;
      R_i[3,17] := -0.23068254;
      R_i[3,18] := -0.28099820;
      R_i[3,19] := -0.18721125;
      R_i[3,20] := -0.10498459;
      R_i[3,21] := -0.46346831;
      R_i[3,22] := -0.27303410;
      R_i[3,23] := -0.16539162;
      R_i[3,24] := 0.75813276;
      R_i[3,25] := -0.42776185;
      R_i[3,26] := 0.37133542;
      R_i[3,27] := 0.56733567;
      R_i[3,28] := -0.40458134;
      R_i[3,29] := 0.52082050;
      R_i[3,30] := -0.03682783;
      R_i[3,31] := -0.11073664;
      R_i[4,0] := -0.27738518;
      R_i[4,1] := 0.21788643;
      R_i[4,2] := -0.03493356;
      R_i[4,3] := -0.38405979;
      R_i[4,4] := -1.14212549;
      R_i[4,5] := -0.69589919;
      R_i[4,6] := -0.48883525;
      R_i[4,7] := -0.06883857;
      R_i[4,8] := 0.19895054;
      R_i[4,9] := 0.14242470;
      R_i[4,10] := -0.35284361;
      R_i[4,11] := -0.20668615;
      R_i[4,12] := -0.09521909;
      R_i[4,13] := -0.30126980;
      R_i[4,14] := -0.29098076;
      R_i[4,15] := 0.26446763;
      R_i[4,16] := -0.12575400;
      R_i[4,17] := 0.08938091;
      R_i[4,18] := 0.21658640;
      R_i[4,19] := -0.36374727;
      R_i[4,20] := -0.52650046;
      R_i[4,21] := -0.61958766;
      R_i[4,22] := -0.55982614;
      R_i[4,23] := 0.45801920;
      R_i[4,24] := -0.62498677;
      R_i[4,25] := 0.59652966;
      R_i[4,26] := 0.50117826;
      R_i[4,27] := -0.26382235;
      R_i[4,28] := 0.31566355;
      R_i[4,29] := 0.17601474;
      R_i[4,30] := 0.37459636;
      R_i[4,31] := 0.24718942;
      R_i[5,0] := -0.26452133;
      R_i[5,1] := -0.45201913;
      R_i[5,2] := 0.05233981;
      R_i[5,3] := 0.34053057;
      R_i[5,4] := 0.29692972;
      R_i[5,5] := -0.74824238;
      R_i[5,6] := 0.11089586;
      R_i[5,7] := -0.27782020;
      R_i[5,8] := -0.15569578;
      R_i[5,9] := 0.18389620;
      R_i[5,10] := 0.01916758;
      R_i[5,11] := -0.12465654;
      R_i[5,12] := -0.11174443;
      R_i[5,13] := 0.02919140;
      R_i[5,14] := -0.47345072;
      R_i[5,15] := 0.13585632;
      R_i[5,16] := -0.05760243;
      R_i[5,17] := 0.41188252;
      R_i[5,18] := 0.19726813;
      R_i[5,19] := 0.02125218;
      R_i[5,20] := -0.02499196;
      R_i[5,21] := 0.05188165;
      R_i[5,22] := 0.01081287;
      R_i[5,23] := -0.02835622;
      R_i[5,24] := -0.05286242;
      R_i[5,25] := 0.05765875;
      R_i[5,26] := 0.09295516;
      R_i[5,27] := 0.26799154;
      R_i[5,28] := -0.39401022;
      R_i[5,29] := 0.50256240;
      R_i[5,30] := -0.20525017;
      R_i[5,31] := -0.12215695;
      R_i[6,0] := -0.20377974;
      R_i[6,1] := 0.45414004;
      R_i[6,2] := -0.15710658;
      R_i[6,3] := -0.34970012;
      R_i[6,4] := -0.02068146;
      R_i[6,5] := -0.10679672;
      R_i[6,6] := -0.38465261;
      R_i[6,7] := 0.01037895;
      R_i[6,8] := 0.29136643;
      R_i[6,9] := 0.28989467;
      R_i[6,10] := -0.37588167;
      R_i[6,11] := -0.16435985;
      R_i[6,12] := -0.35176027;
      R_i[6,13] := 0.23065814;
      R_i[6,14] := -0.16051559;
      R_i[6,15] := -0.09210415;
      R_i[6,16] := -0.11617490;
      R_i[6,17] := 0.33982334;
      R_i[6,18] := 0.08985654;
      R_i[6,19] := -0.17639525;
      R_i[6,20] := 0.36715880;
      R_i[6,21] := 0.16126089;
      R_i[6,22] := 0.06544465;
      R_i[6,23] := -0.30587286;
      R_i[6,24] := 0.12664250;
      R_i[6,25] := 0.22519562;
      R_i[6,26] := 0.14630163;
      R_i[6,27] := -0.09204710;
      R_i[6,28] := 0.23306420;
      R_i[6,29] := -0.14128351;
      R_i[6,30] := -0.01371284;
      R_i[6,31] := -0.58105564;
      R_i[7,0] := -0.05407012;
      R_i[7,1] := -0.22289780;
      R_i[7,2] := -0.00356364;
      R_i[7,3] := -0.33402652;
      R_i[7,4] := 0.48400843;
      R_i[7,5] := 0.16766842;
      R_i[7,6] := 0.04905435;
      R_i[7,7] := 0.30900997;
      R_i[7,8] := -0.21341430;
      R_i[7,9] := 0.05724302;
      R_i[7,10] := -0.23275118;
      R_i[7,11] := -0.29258260;
      R_i[7,12] := 0.33530247;
      R_i[7,13] := -0.07926263;
      R_i[7,14] := -0.61885476;
      R_i[7,15] := 0.11239933;
      R_i[7,16] := -0.65220910;
      R_i[7,17] := 0.25530577;
      R_i[7,18] := -0.09003985;
      R_i[7,19] := -0.31616694;
      R_i[7,20] := -0.02545690;
      R_i[7,21] := 0.05753365;
      R_i[7,22] := 0.29826564;
      R_i[7,23] := -0.27958789;
      R_i[7,24] := 0.25528404;
      R_i[7,25] := -0.44871598;
      R_i[7,26] := 0.16588780;
      R_i[7,27] := -0.31735247;
      R_i[7,28] := -0.27217364;
      R_i[7,29] := -0.06085731;
      R_i[7,30] := -0.13008997;
      R_i[7,31] := -0.13776098;
      R_i[8,0] := -0.35692871;
      R_i[8,1] := 0.04410078;
      R_i[8,2] := -0.44228280;
      R_i[8,3] := 0.01408509;
      R_i[8,4] := 0.36250404;
      R_i[8,5] := 0.06770337;
      R_i[8,6] := -0.18525939;
      R_i[8,7] := -0.17682950;
      R_i[8,8] := -0.25478595;
      R_i[8,9] := 0.08647283;
      R_i[8,10] := 0.48014721;
      R_i[8,11] := 0.02839737;
      R_i[8,12] := 0.10981213;
      R_i[8,13] := 0.01699535;
      R_i[8,14] := 0.19786665;
      R_i[8,15] := -0.03035625;
      R_i[8,16] := -0.31084868;
      R_i[8,17] := -0.18435425;
      R_i[8,18] := 0.33457357;
      R_i[8,19] := -0.22030999;
      R_i[8,20] := 0.12809642;
      R_i[8,21] := -0.27876011;
      R_i[8,22] := 0.00804140;
      R_i[8,23] := -0.15977371;
      R_i[8,24] := 0.19999287;
      R_i[8,25] := -0.03168854;
      R_i[8,26] := 0.01886760;
      R_i[8,27] := -0.17166837;
      R_i[8,28] := -0.13911928;
      R_i[8,29] := 0.17988014;
      R_i[8,30] := 0.01520682;
      R_i[8,31] := 0.14846228;
      R_i[9,0] := -0.41542771;
      R_i[9,1] := 0.20905150;
      R_i[9,2] := 0.23491527;
      R_i[9,3] := -0.21317165;
      R_i[9,4] := 0.34928134;
      R_i[9,5] := 0.25797188;
      R_i[9,6] := 0.15672441;
      R_i[9,7] := 0.02711249;
      R_i[9,8] := -0.10833924;
      R_i[9,9] := 1.00507164;
      R_i[9,10] := 0.18941806;
      R_i[9,11] := -0.57649738;
      R_i[9,12] := -0.10958710;
      R_i[9,13] := -0.27297226;
      R_i[9,14] := -0.11242634;
      R_i[9,15] := 0.07004246;
      R_i[9,16] := -0.49135152;
      R_i[9,17] := 0.33544502;
      R_i[9,18] := 0.34719771;
      R_i[9,19] := 0.20374008;
      R_i[9,20] := 0.00158977;
      R_i[9,21] := -0.13937987;
      R_i[9,22] := 0.33234087;
      R_i[9,23] := -0.08645162;
      R_i[9,24] := 0.05943909;
      R_i[9,25] := 0.03656916;
      R_i[9,26] := 0.21672927;
      R_i[9,27] := -0.02330737;
      R_i[9,28] := -0.10025729;
      R_i[9,29] := 0.14425236;
      R_i[9,30] := -0.03870168;
      R_i[9,31] := -0.04538363;
      R_i[10,0] := 0.36769497;
      R_i[10,1] := 0.09163627;
      R_i[10,2] := 0.01542166;
      R_i[10,3] := -0.08378920;
      R_i[10,4] := 0.50972462;
      R_i[10,5] := -0.16758412;
      R_i[10,6] := 0.04439653;
      R_i[10,7] := 0.17410386;
      R_i[10,8] := -0.23226380;
      R_i[10,9] := 0.19068857;
      R_i[10,10] := -0.42978424;
      R_i[10,11] := -0.02443463;
      R_i[10,12] := 0.17334399;
      R_i[10,13] := 0.14308771;
      R_i[10,14] := 0.42658469;
      R_i[10,15] := 0.08669236;
      R_i[10,16] := -0.14037156;
      R_i[10,17] := 0.15868302;
      R_i[10,18] := 0.10887319;
      R_i[10,19] := 0.01519258;
      R_i[10,20] := 0.09982713;
      R_i[10,21] := -0.13058648;
      R_i[10,22] := 0.06128490;
      R_i[10,23] := 0.09715474;
      R_i[10,24] := 0.01161596;
      R_i[10,25] := 0.00869740;
      R_i[10,26] := 0.15081570;
      R_i[10,27] := -0.40050906;
      R_i[10,28] := 0.07687394;
      R_i[10,29] := -0.18552521;
      R_i[10,30] := -0.02003719;
      R_i[10,31] := 0.08377120;
      R_i[11,0] := -0.01316699;
      R_i[11,1] := 0.10122313;
      R_i[11,2] := -0.10969920;
      R_i[11,3] := -0.23030835;
      R_i[11,4] := 0.60010606;
      R_i[11,5] := -0.34940866;
      R_i[11,6] := 0.31191304;
      R_i[11,7] := 0.31473544;
      R_i[11,8] := 0.12409268;
      R_i[11,9] := -0.00975981;
      R_i[11,10] := 0.36657432;
      R_i[11,11] := 1.10749483;
      R_i[11,12] := 0.01427285;
      R_i[11,13] := 0.28292170;
      R_i[11,14] := -0.73101860;
      R_i[11,15] := -0.17629677;
      R_i[11,16] := -0.24775396;
      R_i[11,17] := -0.17321597;
      R_i[11,18] := -0.28576198;
      R_i[11,19] := -0.16400611;
      R_i[11,20] := 0.58374870;
      R_i[11,21] := -0.23495102;
      R_i[11,22] := 0.67055702;
      R_i[11,23] := -0.64832348;
      R_i[11,24] := 0.41382262;
      R_i[11,25] := -0.56086731;
      R_i[11,26] := -0.37854087;
      R_i[11,27] := -0.33385524;
      R_i[11,28] := 0.35420173;
      R_i[11,29] := 0.09360323;
      R_i[11,30] := -0.12521435;
      R_i[11,31] := -0.70395684;
      R_i[12,0] := -0.34958652;
      R_i[12,1] := -0.04477185;
      R_i[12,2] := 0.17206842;
      R_i[12,3] := 0.33812946;
      R_i[12,4] := -0.16370592;
      R_i[12,5] := 0.35788283;
      R_i[12,6] := 0.25873747;
      R_i[12,7] := -0.25274616;
      R_i[12,8] := -0.31537613;
      R_i[12,9] := -0.10520653;
      R_i[12,10] := 0.27170977;
      R_i[12,11] := 0.03155406;
      R_i[12,12] := 0.61352289;
      R_i[12,13] := -0.11578090;
      R_i[12,14] := 0.06411036;
      R_i[12,15] := -0.06842072;
      R_i[12,16] := -0.03340700;
      R_i[12,17] := 0.17851020;
      R_i[12,18] := 0.05276991;
      R_i[12,19] := -0.27957132;
      R_i[12,20] := 0.09669928;
      R_i[12,21] := -0.25238210;
      R_i[12,22] := 0.24651983;
      R_i[12,23] := -0.18397731;
      R_i[12,24] := 0.02993304;
      R_i[12,25] := 0.18756384;
      R_i[12,26] := 0.03975990;
      R_i[12,27] := -0.22840789;
      R_i[12,28] := 0.23632295;
      R_i[12,29] := 0.15286604;
      R_i[12,30] := -0.09223666;
      R_i[12,31] := 0.11066151;
      R_i[13,0] := -0.18651058;
      R_i[13,1] := 0.21643525;
      R_i[13,2] := 0.12474846;
      R_i[13,3] := 0.09924160;
      R_i[13,4] := -0.06626517;
      R_i[13,5] := 0.07129208;
      R_i[13,6] := -0.60450929;
      R_i[13,7] := -0.08253109;
      R_i[13,8] := 0.11061417;
      R_i[13,9] := -0.14199089;
      R_i[13,10] := -0.00901213;
      R_i[13,11] := 0.01251668;
      R_i[13,12] := 0.40270495;
      R_i[13,13] := 0.16962376;
      R_i[13,14] := -0.31417164;
      R_i[13,15] := -0.13672313;
      R_i[13,16] := 0.42094859;
      R_i[13,17] := -0.31583846;
      R_i[13,18] := -0.19630848;
      R_i[13,19] := -0.23622292;
      R_i[13,20] := 0.11617036;
      R_i[13,21] := -0.48445079;
      R_i[13,22] := -0.46077368;
      R_i[13,23] := -0.10126588;
      R_i[13,24] := 0.08009661;
      R_i[13,25] := 0.09753137;
      R_i[13,26] := -0.02010051;
      R_i[13,27] := -0.12881830;
      R_i[13,28] := 0.23913288;
      R_i[13,29] := -0.37161407;
      R_i[13,30] := 0.21826558;
      R_i[13,31] := 0.23566197;
      R_i[14,0] := -0.22003971;
      R_i[14,1] := 0.11151226;
      R_i[14,2] := 0.11048436;
      R_i[14,3] := 0.15629630;
      R_i[14,4] := 0.06400732;
      R_i[14,5] := 0.32734475;
      R_i[14,6] := -0.03265190;
      R_i[14,7] := -0.25161412;
      R_i[14,8] := -0.04165458;
      R_i[14,9] := 0.27729705;
      R_i[14,10] := 0.82511091;
      R_i[14,11] := -0.30799398;
      R_i[14,12] := -0.01025582;
      R_i[14,13] := -0.11674581;
      R_i[14,14] := -2.80562019;
      R_i[14,15] := 0.52282768;
      R_i[14,16] := -0.09129780;
      R_i[14,17] := -0.00227208;
      R_i[14,18] := 0.39883411;
      R_i[14,19] := -0.16658033;
      R_i[14,20] := -0.07539129;
      R_i[14,21] := 0.15584196;
      R_i[14,22] := -0.00372907;
      R_i[14,23] := 0.14898381;
      R_i[14,24] := 0.15867527;
      R_i[14,25] := 0.13778594;
      R_i[14,26] := 0.16674924;
      R_i[14,27] := 0.41589451;
      R_i[14,28] := -0.16052705;
      R_i[14,29] := 0.06137883;
      R_i[14,30] := 0.17442019;
      R_i[14,31] := 0.01023346;
      R_i[15,0] := 0.49395472;
      R_i[15,1] := 0.19703144;
      R_i[15,2] := -0.08435930;
      R_i[15,3] := 0.34724095;
      R_i[15,4] := 0.29099765;
      R_i[15,5] := -0.24459985;
      R_i[15,6] := 0.26904958;
      R_i[15,7] := -0.20164552;
      R_i[15,8] := -0.24098852;
      R_i[15,9] := -0.18421091;
      R_i[15,10] := 0.00619574;
      R_i[15,11] := 0.26867259;
      R_i[15,12] := -0.17595857;
      R_i[15,13] := -0.05126722;
      R_i[15,14] := -0.09862539;
      R_i[15,15] := 0.68389630;
      R_i[15,16] := -0.18652491;
      R_i[15,17] := 0.02966011;
      R_i[15,18] := -0.25917655;
      R_i[15,19] := 0.04642781;
      R_i[15,20] := 0.00999165;
      R_i[15,21] := 0.38628080;
      R_i[15,22] := -0.06190461;
      R_i[15,23] := -0.03847435;
      R_i[15,24] := -0.25492656;
      R_i[15,25] := -0.08687152;
      R_i[15,26] := 0.49867639;
      R_i[15,27] := -0.20988461;
      R_i[15,28] := 0.20958014;
      R_i[15,29] := 0.02616844;
      R_i[15,30] := -0.19732095;
      R_i[15,31] := -0.20276946;
      R_i[16,0] := -0.19701254;
      R_i[16,1] := 0.03600208;
      R_i[16,2] := 0.13406947;
      R_i[16,3] := -0.06813481;
      R_i[16,4] := -0.01291389;
      R_i[16,5] := 0.49659860;
      R_i[16,6] := 0.10141860;
      R_i[16,7] := -0.91545212;
      R_i[16,8] := -1.25405025;
      R_i[16,9] := 0.11031634;
      R_i[16,10] := -0.10669987;
      R_i[16,11] := 0.24751085;
      R_i[16,12] := -0.21095966;
      R_i[16,13] := -0.23712406;
      R_i[16,14] := -0.22438581;
      R_i[16,15] := 0.33338776;
      R_i[16,16] := -0.47963321;
      R_i[16,17] := -0.23448418;
      R_i[16,18] := -0.21523100;
      R_i[16,19] := 0.10917976;
      R_i[16,20] := -0.01618838;
      R_i[16,21] := 0.12323362;
      R_i[16,22] := -0.43334574;
      R_i[16,23] := 0.30341670;
      R_i[16,24] := 0.28056833;
      R_i[16,25] := 0.47891304;
      R_i[16,26] := 0.04055469;
      R_i[16,27] := -0.04559619;
      R_i[16,28] := 0.26704851;
      R_i[16,29] := 0.19118740;
      R_i[16,30] := -0.38988611;
      R_i[16,31] := 0.05536282;
      R_i[17,0] := -0.25103343;
      R_i[17,1] := 0.00119750;
      R_i[17,2] := -0.32162443;
      R_i[17,3] := -0.42256883;
      R_i[17,4] := 0.05387824;
      R_i[17,5] := -0.01850677;
      R_i[17,6] := 0.16165783;
      R_i[17,7] := -0.18163699;
      R_i[17,8] := -0.14975813;
      R_i[17,9] := 0.53523248;
      R_i[17,10] := 0.44817653;
      R_i[17,11] := -0.58926225;
      R_i[17,12] := -0.28382024;
      R_i[17,13] := -0.32453334;
      R_i[17,14] := -0.00467656;
      R_i[17,15] := 0.07768948;
      R_i[17,16] := -0.82502997;
      R_i[17,17] := 1.91944230;
      R_i[17,18] := 0.43120643;
      R_i[17,19] := 0.10850436;
      R_i[17,20] := 0.01053265;
      R_i[17,21] := -0.07928012;
      R_i[17,22] := 0.02779940;
      R_i[17,23] := -0.04494777;
      R_i[17,24] := 0.02061015;
      R_i[17,25] := 0.19665171;
      R_i[17,26] := 0.36106840;
      R_i[17,27] := -0.06449664;
      R_i[17,28] := -0.20015582;
      R_i[17,29] := 0.18195516;
      R_i[17,30] := -0.10667004;
      R_i[17,31] := -0.16377114;
      R_i[18,0] := 0.14792579;
      R_i[18,1] := -0.23028043;
      R_i[18,2] := 0.06688867;
      R_i[18,3] := -0.95816082;
      R_i[18,4] := -0.17983703;
      R_i[18,5] := -0.14859901;
      R_i[18,6] := 0.05815475;
      R_i[18,7] := -0.46422938;
      R_i[18,8] := 0.33274713;
      R_i[18,9] := 0.08284145;
      R_i[18,10] := -0.56101692;
      R_i[18,11] := -0.64956868;
      R_i[18,12] := -0.51611423;
      R_i[18,13] := -0.08295774;
      R_i[18,14] := -0.71968442;
      R_i[18,15] := 0.65384507;
      R_i[18,16] := -0.42235219;
      R_i[18,17] := 0.61090374;
      R_i[18,18] := 0.10827148;
      R_i[18,19] := -0.52440095;
      R_i[18,20] := -0.30586541;
      R_i[18,21] := 0.19868562;
      R_i[18,22] := 0.47836059;
      R_i[18,23] := 0.17784643;
      R_i[18,24] := -0.56319577;
      R_i[18,25] := 0.21957074;
      R_i[18,26] := -0.19798693;
      R_i[18,27] := 0.15806785;
      R_i[18,28] := -0.24106851;
      R_i[18,29] := 0.02314841;
      R_i[18,30] := -0.05501189;
      R_i[18,31] := -0.39892396;
      R_i[19,0] := 0.16951925;
      R_i[19,1] := 0.25170106;
      R_i[19,2] := 0.04045393;
      R_i[19,3] := -0.47197193;
      R_i[19,4] := -0.30712649;
      R_i[19,5] := -0.02992622;
      R_i[19,6] := 0.14370751;
      R_i[19,7] := -0.06286702;
      R_i[19,8] := 0.23131999;
      R_i[19,9] := 0.15838535;
      R_i[19,10] := 1.18502522;
      R_i[19,11] := 0.12588599;
      R_i[19,12] := -0.21159452;
      R_i[19,13] := 0.03646610;
      R_i[19,14] := 0.05060637;
      R_i[19,15] := 0.25694394;
      R_i[19,16] := -0.70235902;
      R_i[19,17] := 0.06837672;
      R_i[19,18] := 0.17778705;
      R_i[19,19] := -1.18717599;
      R_i[19,20] := -0.06324542;
      R_i[19,21] := -0.38142931;
      R_i[19,22] := -0.71301126;
      R_i[19,23] := 0.27857348;
      R_i[19,24] := -0.42894375;
      R_i[19,25] := 0.04813502;
      R_i[19,26] := 0.11246923;
      R_i[19,27] := -0.35118386;
      R_i[19,28] := -0.39048925;
      R_i[19,29] := 0.37312102;
      R_i[19,30] := -0.33647817;
      R_i[19,31] := 0.53995860;
      R_i[20,0] := 0.25687960;
      R_i[20,1] := -0.29242688;
      R_i[20,2] := 0.37741703;
      R_i[20,3] := 0.30777171;
      R_i[20,4] := -0.20866543;
      R_i[20,5] := -0.01098926;
      R_i[20,6] := 0.11667342;
      R_i[20,7] := -0.55857700;
      R_i[20,8] := -0.05032220;
      R_i[20,9] := -0.04135040;
      R_i[20,10] := 0.51183265;
      R_i[20,11] := -0.49198973;
      R_i[20,12] := -0.34401676;
      R_i[20,13] := -0.02927491;
      R_i[20,14] := -0.17992254;
      R_i[20,15] := -0.38016060;
      R_i[20,16] := -0.38633218;
      R_i[20,17] := 0.59576029;
      R_i[20,18] := 0.34693968;
      R_i[20,19] := 0.11619298;
      R_i[20,20] := -0.26961488;
      R_i[20,21] := -0.47565496;
      R_i[20,22] := 0.14985557;
      R_i[20,23] := -0.01094213;
      R_i[20,24] := -0.08863560;
      R_i[20,25] := -0.13210621;
      R_i[20,26] := 0.17917508;
      R_i[20,27] := 0.09925277;
      R_i[20,28] := 0.30064869;
      R_i[20,29] := -0.60817754;
      R_i[20,30] := -0.18754429;
      R_i[20,31] := -0.24060634;
      R_i[21,0] := 0.08565907;
      R_i[21,1] := -0.44212258;
      R_i[21,2] := -0.91510022;
      R_i[21,3] := 0.21750584;
      R_i[21,4] := -0.20699133;
      R_i[21,5] := 0.12427791;
      R_i[21,6] := -0.79080284;
      R_i[21,7] := -0.01921312;
      R_i[21,8] := -0.92770261;
      R_i[21,9] := -0.12546726;
      R_i[21,10] := -0.80846310;
      R_i[21,11] := -0.09977988;
      R_i[21,12] := -1.13460350;
      R_i[21,13] := 0.02645151;
      R_i[21,14] := -0.92707533;
      R_i[21,15] := -0.44168460;
      R_i[21,16] := -0.57176465;
      R_i[21,17] := 0.39779779;
      R_i[21,18] := -0.12863410;
      R_i[21,19] := 0.54696029;
      R_i[21,20] := -1.60230041;
      R_i[21,21] := -3.06046152;
      R_i[21,22] := 0.87443531;
      R_i[21,23] := -0.35160878;
      R_i[21,24] := 0.45174626;
      R_i[21,25] := 0.65975076;
      R_i[21,26] := 0.43925485;
      R_i[21,27] := 0.15303802;
      R_i[21,28] := 0.55273247;
      R_i[21,29] := 0.91924977;
      R_i[21,30] := 0.57290447;
      R_i[21,31] := -0.41661522;
      R_i[22,0] := 0.23858294;
      R_i[22,1] := 0.30541795;
      R_i[22,2] := 0.09449539;
      R_i[22,3] := -0.42065448;
      R_i[22,4] := -0.16242130;
      R_i[22,5] := -0.24975078;
      R_i[22,6] := -0.01201073;
      R_i[22,7] := -0.59941405;
      R_i[22,8] := -0.18639621;
      R_i[22,9] := 0.28788194;
      R_i[22,10] := -0.56155074;
      R_i[22,11] := 0.41028517;
      R_i[22,12] := 0.07601306;
      R_i[22,13] := 0.00874536;
      R_i[22,14] := -0.26729393;
      R_i[22,15] := 0.28428996;
      R_i[22,16] := -0.51269424;
      R_i[22,17] := 0.05877603;
      R_i[22,18] := 0.40804940;
      R_i[22,19] := -0.08256710;
      R_i[22,20] := -0.01787679;
      R_i[22,21] := 0.07941986;
      R_i[22,22] := 0.51579964;
      R_i[22,23] := 0.06920873;
      R_i[22,24] := 0.07815367;
      R_i[22,25] := 0.09119307;
      R_i[22,26] := 0.26356244;
      R_i[22,27] := 0.03236705;
      R_i[22,28] := 0.41603360;
      R_i[22,29] := -0.23240425;
      R_i[22,30] := -0.49368262;
      R_i[22,31] := -0.23237231;
      R_i[23,0] := -0.11686549;
      R_i[23,1] := 0.59647936;
      R_i[23,2] := -0.09401071;
      R_i[23,3] := -0.17464159;
      R_i[23,4] := 0.56050313;
      R_i[23,5] := -0.10255875;
      R_i[23,6] := 0.47642258;
      R_i[23,7] := 0.03974510;
      R_i[23,8] := -0.30848908;
      R_i[23,9] := -0.08085486;
      R_i[23,10] := 0.10946240;
      R_i[23,11] := -0.03398137;
      R_i[23,12] := -0.23338807;
      R_i[23,13] := -0.38847858;
      R_i[23,14] := 0.12661757;
      R_i[23,15] := -0.13903099;
      R_i[23,16] := -0.54911894;
      R_i[23,17] := 0.05592053;
      R_i[23,18] := -0.06480610;
      R_i[23,19] := -0.40487275;
      R_i[23,20] := 0.35428700;
      R_i[23,21] := 0.13950250;
      R_i[23,22] := 0.51759350;
      R_i[23,23] := 0.79979062;
      R_i[23,24] := 0.67532921;
      R_i[23,25] := -0.35276383;
      R_i[23,26] := 0.26916650;
      R_i[23,27] := -0.22992319;
      R_i[23,28] := 0.37736148;
      R_i[23,29] := 0.22526073;
      R_i[23,30] := 0.19747670;
      R_i[23,31] := -0.94982904;
      R_i[24,0] := 0.11757268;
      R_i[24,1] := 0.26305696;
      R_i[24,2] := -0.23278375;
      R_i[24,3] := -0.06885347;
      R_i[24,4] := -0.11244328;
      R_i[24,5] := -0.46475348;
      R_i[24,6] := -0.37523627;
      R_i[24,7] := -0.18539278;
      R_i[24,8] := 0.13196871;
      R_i[24,9] := -0.26032043;
      R_i[24,10] := -0.35013422;
      R_i[24,11] := 0.25641710;
      R_i[24,12] := -0.11111728;
      R_i[24,13] := 0.22136630;
      R_i[24,14] := -0.19546731;
      R_i[24,15] := -0.08531215;
      R_i[24,16] := 0.10026735;
      R_i[24,17] := -0.44211304;
      R_i[24,18] := -0.10861719;
      R_i[24,19] := -0.29563421;
      R_i[24,20] := -0.12760343;
      R_i[24,21] := 0.06214319;
      R_i[24,22] := -0.39911950;
      R_i[24,23] := 0.27528340;
      R_i[24,24] := -0.33778524;
      R_i[24,25] := -0.02838964;
      R_i[24,26] := 0.36320505;
      R_i[24,27] := -0.33704430;
      R_i[24,28] := 0.08388724;
      R_i[24,29] := 0.06718535;
      R_i[24,30] := -0.10252665;
      R_i[24,31] := -0.14726697;
      R_i[25,0] := -0.31382275;
      R_i[25,1] := 0.15260525;
      R_i[25,2] := -0.26525092;
      R_i[25,3] := -0.01837087;
      R_i[25,4] := 0.50268316;
      R_i[25,5] := 0.28868583;
      R_i[25,6] := -0.21333495;
      R_i[25,7] := 0.05177091;
      R_i[25,8] := -0.55214375;
      R_i[25,9] := 0.33633831;
      R_i[25,10] := 0.19150658;
      R_i[25,11] := -0.53368002;
      R_i[25,12] := 0.25028932;
      R_i[25,13] := 0.32556430;
      R_i[25,14] := -0.25146353;
      R_i[25,15] := 0.15585208;
      R_i[25,16] := -0.50763589;
      R_i[25,17] := 0.60535324;
      R_i[25,18] := 0.16541542;
      R_i[25,19] := -0.04087145;
      R_i[25,20] := 0.04982444;
      R_i[25,21] := -0.18684447;
      R_i[25,22] := 0.34545532;
      R_i[25,23] := 0.01859861;
      R_i[25,24] := 0.36723447;
      R_i[25,25] := 0.02203113;
      R_i[25,26] := 0.21915229;
      R_i[25,27] := -0.12987208;
      R_i[25,28] := -0.06913047;
      R_i[25,29] := -0.18187772;
      R_i[25,30] := -0.20342335;
      R_i[25,31] := -0.10493086;
      R_i[26,0] := -0.53719932;
      R_i[26,1] := -0.13339937;
      R_i[26,2] := 0.05625769;
      R_i[26,3] := -0.38640153;
      R_i[26,4] := -0.50864387;
      R_i[26,5] := 0.31767592;
      R_i[26,6] := -0.05330179;
      R_i[26,7] := -0.18287997;
      R_i[26,8] := -0.55325216;
      R_i[26,9] := 0.04128635;
      R_i[26,10] := 0.23983631;
      R_i[26,11] := -0.71368462;
      R_i[26,12] := -0.17042463;
      R_i[26,13] := -0.17299728;
      R_i[26,14] := -0.63668227;
      R_i[26,15] := 1.12886727;
      R_i[26,16] := -0.69215649;
      R_i[26,17] := 0.14695346;
      R_i[26,18] := 0.02460258;
      R_i[26,19] := -0.11582782;
      R_i[26,20] := 0.14957139;
      R_i[26,21] := -1.03943086;
      R_i[26,22] := -0.04483403;
      R_i[26,23] := -0.13662077;
      R_i[26,24] := -0.10242261;
      R_i[26,25] := 0.01423822;
      R_i[26,26] := -1.68651748;
      R_i[26,27] := 0.28457990;
      R_i[26,28] := -0.05783774;
      R_i[26,29] := 0.91989142;
      R_i[26,30] := 0.84364921;
      R_i[26,31] := -0.14265282;
      R_i[27,0] := -0.01278794;
      R_i[27,1] := 0.64636630;
      R_i[27,2] := 0.05488608;
      R_i[27,3] := -0.04217035;
      R_i[27,4] := 0.43805686;
      R_i[27,5] := 0.29401278;
      R_i[27,6] := 0.05735238;
      R_i[27,7] := 0.24532473;
      R_i[27,8] := 0.09328273;
      R_i[27,9] := 0.20191593;
      R_i[27,10] := -0.05074343;
      R_i[27,11] := -0.07691138;
      R_i[27,12] := -0.10834948;
      R_i[27,13] := -0.32525727;
      R_i[27,14] := -0.27253160;
      R_i[27,15] := -0.25859049;
      R_i[27,16] := -0.14507720;
      R_i[27,17] := 0.28425568;
      R_i[27,18] := 0.37385944;
      R_i[27,19] := 0.26338044;
      R_i[27,20] := 0.56770164;
      R_i[27,21] := 0.03139745;
      R_i[27,22] := 0.16119128;
      R_i[27,23] := -0.31055555;
      R_i[27,24] := 0.13619593;
      R_i[27,25] := -0.18741760;
      R_i[27,26] := 0.16516344;
      R_i[27,27] := 0.24178873;
      R_i[27,28] := -0.12709211;
      R_i[27,29] := 0.08763196;
      R_i[27,30] := -0.14837472;
      R_i[27,31] := -0.32929465;
      R_i[28,0] := -0.04833423;
      R_i[28,1] := -0.06972695;
      R_i[28,2] := 0.12358193;
      R_i[28,3] := -0.00748151;
      R_i[28,4] := 0.20087366;
      R_i[28,5] := 0.02704377;
      R_i[28,6] := 0.31676322;
      R_i[28,7] := -0.08208895;
      R_i[28,8] := 0.70627993;
      R_i[28,9] := -0.41975358;
      R_i[28,10] := -0.03168092;
      R_i[28,11] := -0.24489982;
      R_i[28,12] := 0.01355535;
      R_i[28,13] := -0.02193020;
      R_i[28,14] := 0.39523152;
      R_i[28,15] := -0.07223310;
      R_i[28,16] := -0.02367456;
      R_i[28,17] := 0.55328524;
      R_i[28,18] := -0.34179929;
      R_i[28,19] := -0.36209509;
      R_i[28,20] := 0.14367893;
      R_i[28,21] := -0.50094742;
      R_i[28,22] := -0.24588630;
      R_i[28,23] := -0.01608187;
      R_i[28,24] := 0.05603309;
      R_i[28,25] := -0.30418012;
      R_i[28,26] := 0.14532541;
      R_i[28,27] := -0.02157391;
      R_i[28,28] := 0.43848851;
      R_i[28,29] := 0.26743150;
      R_i[28,30] := -0.39355049;
      R_i[28,31] := -0.42640853;
      R_i[29,0] := -0.19193545;
      R_i[29,1] := -0.37056381;
      R_i[29,2] := -0.36622241;
      R_i[29,3] := -0.13623630;
      R_i[29,4] := 0.12658711;
      R_i[29,5] := 0.43985888;
      R_i[29,6] := 0.00195898;
      R_i[29,7] := 0.03340083;
      R_i[29,8] := 0.01248389;
      R_i[29,9] := -0.18806490;
      R_i[29,10] := -0.34636173;
      R_i[29,11] := -0.26499057;
      R_i[29,12] := 0.22303945;
      R_i[29,13] := -1.19130385;
      R_i[29,14] := 0.50972050;
      R_i[29,15] := 0.55376738;
      R_i[29,16] := 0.25370732;
      R_i[29,17] := 0.05993506;
      R_i[29,18] := 0.05035046;
      R_i[29,19] := 0.36397049;
      R_i[29,20] := -0.26611117;
      R_i[29,21] := -0.30689833;
      R_i[29,22] := 1.33433664;
      R_i[29,23] := -0.36145219;
      R_i[29,24] := -0.64593756;
      R_i[29,25] := -0.04382587;
      R_i[29,26] := 0.90402567;
      R_i[29,27] := -0.08520819;
      R_i[29,28] := -1.02085721;
      R_i[29,29] := -4.01971674;
      R_i[29,30] := -0.36914620;
      R_i[29,31] := -0.78251827;
      R_i[30,0] := -0.16355217;
      R_i[30,1] := 0.39272520;
      R_i[30,2] := -0.59471846;
      R_i[30,3] := -0.14043310;
      R_i[30,4] := 0.32514334;
      R_i[30,5] := 0.29283226;
      R_i[30,6] := 0.62080425;
      R_i[30,7] := -0.49486405;
      R_i[30,8] := -0.21475920;
      R_i[30,9] := 1.07951474;
      R_i[30,10] := 0.85024750;
      R_i[30,11] := -0.21696174;
      R_i[30,12] := 0.32457268;
      R_i[30,13] := -0.29199421;
      R_i[30,14] := 0.00222744;
      R_i[30,15] := -0.24674690;
      R_i[30,16] := -0.27139488;
      R_i[30,17] := 0.03089927;
      R_i[30,18] := 0.17938614;
      R_i[30,19] := -0.48254132;
      R_i[30,20] := 0.20032924;
      R_i[30,21] := -0.03424564;
      R_i[30,22] := 0.98936754;
      R_i[30,23] := -0.56116986;
      R_i[30,24] := 0.13367562;
      R_i[30,25] := 0.74008280;
      R_i[30,26] := -0.02666840;
      R_i[30,27] := 0.04185103;
      R_i[30,28] := 0.45641306;
      R_i[30,29] := -0.16268258;
      R_i[30,30] := 2.80819917;
      R_i[30,31] := -1.14883232;
      R_i[31,0] := -0.11986776;
      R_i[31,1] := -0.48983297;
      R_i[31,2] := -0.25225723;
      R_i[31,3] := 0.23466448;
      R_i[31,4] := 0.37974370;
      R_i[31,5] := -0.02909207;
      R_i[31,6] := 0.34044248;
      R_i[31,7] := 0.36115289;
      R_i[31,8] := 0.06270733;
      R_i[31,9] := -0.33002385;
      R_i[31,10] := 0.04319567;
      R_i[31,11] := -0.65197051;
      R_i[31,12] := -0.13991827;
      R_i[31,13] := -0.51894534;
      R_i[31,14] := -0.19465037;
      R_i[31,15] := 0.09193419;
      R_i[31,16] := -0.46575260;
      R_i[31,17] := 0.81263840;
      R_i[31,18] := -0.02694119;
      R_i[31,19] := -0.62276167;
      R_i[31,20] := 0.23468377;
      R_i[31,21] := -0.18955506;
      R_i[31,22] := 0.13500233;
      R_i[31,23] := 0.04741247;
      R_i[31,24] := -0.00523690;
      R_i[31,25] := -0.40990052;
      R_i[31,26] := -0.05144414;
      R_i[31,27] := -0.27209201;
      R_i[31,28] := 0.06281765;
      R_i[31,29] := 0.50419718;
      R_i[31,30] := -0.00771237;
      R_i[31,31] := 0.04130097;
      R_f[0,0] := -0.67533004;
      R_f[0,1] := 0.02714094;
      R_f[0,2] := -0.43118471;
      R_f[0,3] := -0.24901403;
      R_f[0,4] := -0.28021365;
      R_f[0,5] := -0.22351769;
      R_f[0,6] := -0.09202358;
      R_f[0,7] := -0.35974187;
      R_f[0,8] := 0.04250066;
      R_f[0,9] := -0.70527303;
      R_f[0,10] := 0.64902079;
      R_f[0,11] := -0.80287552;
      R_f[0,12] := -0.62369150;
      R_f[0,13] := 0.01997556;
      R_f[0,14] := 0.33401716;
      R_f[0,15] := -0.02997861;
      R_f[0,16] := 0.16724707;
      R_f[0,17] := -0.09938758;
      R_f[0,18] := 0.12572917;
      R_f[0,19] := -0.22990333;
      R_f[0,20] := -0.35627905;
      R_f[0,21] := -0.66718334;
      R_f[0,22] := 0.64487123;
      R_f[0,23] := -0.39761934;
      R_f[0,24] := 0.11252652;
      R_f[0,25] := 0.35531715;
      R_f[0,26] := -0.12102325;
      R_f[0,27] := 0.06884732;
      R_f[0,28] := -0.35347942;
      R_f[0,29] := -0.66960865;
      R_f[0,30] := 0.37912908;
      R_f[0,31] := 0.14283381;
      R_f[1,0] := 0.48609182;
      R_f[1,1] := 0.61146563;
      R_f[1,2] := -0.36975044;
      R_f[1,3] := 0.50827461;
      R_f[1,4] := 0.09001865;
      R_f[1,5] := -0.33936116;
      R_f[1,6] := 0.35342741;
      R_f[1,7] := 0.25101903;
      R_f[1,8] := -0.44604495;
      R_f[1,9] := -0.13113552;
      R_f[1,10] := 0.71121246;
      R_f[1,11] := -0.71102190;
      R_f[1,12] := -0.66324550;
      R_f[1,13] := -0.44045416;
      R_f[1,14] := -0.61123687;
      R_f[1,15] := 0.35812396;
      R_f[1,16] := 0.04237995;
      R_f[1,17] := -0.53959906;
      R_f[1,18] := 0.82591206;
      R_f[1,19] := 0.03209597;
      R_f[1,20] := 0.41162083;
      R_f[1,21] := 0.77022076;
      R_f[1,22] := 0.11187772;
      R_f[1,23] := -0.04342550;
      R_f[1,24] := 0.43034852;
      R_f[1,25] := -0.07955813;
      R_f[1,26] := 0.52373642;
      R_f[1,27] := 0.25399476;
      R_f[1,28] := 0.27276284;
      R_f[1,29] := -0.93637961;
      R_f[1,30] := 0.06395336;
      R_f[1,31] := 0.05123950;
      R_f[2,0] := -0.05785920;
      R_f[2,1] := -0.00636479;
      R_f[2,2] := -0.55666709;
      R_f[2,3] := -0.53078192;
      R_f[2,4] := 0.61353374;
      R_f[2,5] := -0.76166481;
      R_f[2,6] := -0.13201754;
      R_f[2,7] := 0.63591111;
      R_f[2,8] := 0.68129236;
      R_f[2,9] := -0.83181989;
      R_f[2,10] := 0.26337647;
      R_f[2,11] := 0.02993034;
      R_f[2,12] := -1.28638637;
      R_f[2,13] := -0.45174307;
      R_f[2,14] := 0.46492049;
      R_f[2,15] := 0.28912774;
      R_f[2,16] := 0.80125827;
      R_f[2,17] := -0.66417259;
      R_f[2,18] := 0.37046370;
      R_f[2,19] := -0.98936939;
      R_f[2,20] := 0.02043331;
      R_f[2,21] := -0.84147042;
      R_f[2,22] := 0.42977002;
      R_f[2,23] := -0.45103595;
      R_f[2,24] := 0.52417392;
      R_f[2,25] := -0.32892042;
      R_f[2,26] := -0.01681360;
      R_f[2,27] := -0.65100932;
      R_f[2,28] := -0.02503461;
      R_f[2,29] := -0.27034515;
      R_f[2,30] := -0.09233637;
      R_f[2,31] := 0.09730685;
